(* IEC 61131-3 sources: daoli-st-library/DL_Algo (part 2) *)

(* ---- FB_DL_LuenbergerObserver.st ---- *)
(*==============================================================================
 * 组件名称 (Component)  : FB_DL_LuenbergerObserver
 * 所属子库 (Sublibrary) : DL_Algo
 * 当前版本 (Version)    : 1.0.1
 * 兼容性   (Platform)   : CODESYS 3.5+ / TwinCAT 3 / 汇川 InoProShop / 施耐德 Machine Expert
 *                         仅依赖 Standard.library（TON / R_TRIG / ABS / SQRT / MIN / MAX），零厂商私有库
 * 功能描述 (Function)   : 离散二阶状态观测器（Luenberger 结构）+ 残差窗收敛判据 + 防发散钳位。
 *                         被估对象为二阶线性离散模型（位置/速度）：
 *                           x1⁺ = a11·x1 + a12·x2 + b1·u        （位置方程）
 *                           x2⁺ = a21·x1 + a22·x2 + b2·u        （速度方程）
 *                           yHat = x1⁺                           （测点为位置）
 *                         观测器（Luenberger 增益 L = [l1, l2]）：
 *                           r  = y − yHat（新息）
 *                           x1 = x1⁺ + l1·r
 *                           x2 = x2⁺ + l2·r
 *                         收敛判据：以周期窗（自复位 TON）为单位累计新息平方和，窗末算均方根
 *                         fResRms = SQRT(Σr²/n)。fResRms <= fResThr 记为收敛（bConverged 置真），
 *                         否则清零。**只有收敛后才宣称状态估计可用**——不收敛时 x1Hat/x2Hat 仍输出
 *                         （便于诊断），但 bEstValid=FALSE，不得参与闭环。
 *                         防发散：① 每个状态在更新后钳到 ±fXMax，触位即 bClamped（饱和非故障）；
 *                         ② 窗 RMS 超 fResDiv 判观测器发散（故障锁存，eCause=eDiverged），
 *                         因为真实系统残差不会长期比噪声大一个量级；③ 增益/系数 NaN 一律闸死。
 * 接口     (Interface)  : 输入 fY 实测位置、fU 控制量、六个模型系数（a11/a12/a21/a22/b1/b2）、
 *                         两个增益（l1/l2）、fXMax 状态硬限、fResThr 收敛阈、fResDiv 发散阈、
 *                         tWindow 残差窗、bReset；输出 fX1Hat / fX2Hat 状态估计、fResidual 当拍新息、
 *                         fResRms 窗均方根、bConverged 收敛、bEstValid 估计可用、bClamped 触限、
 *                         eState / eCause / bError。
 * 边界     (Boundary)   : ① **属主边界（写死）：本件是纯算法件——不读轴接口、不发指令、
 *                         不参与闭环**。估计值经上层注入，是否用于前馈/诊断由上层决定。
 *                         ② 模型系数与增益由调用方给（本件不做模型辨识）：辨识属 `FB_DL_RlsEstimator`；
 *                         二者可级联（辨识出系数喂本件），但不得互相内嵌。
 *                         ③ 组态闸：fXMax <= DL_LUO_EPS、fResThr <= 0.0、fResDiv <= fResThr、
 *                         tWindow <= T#0S、任一系数/增益/引脚 NaN → 故障锁存，估计输出置 0
 *                         （安全侧：不宣称任何状态）。
 *                         ④ 周期窗用 IN := (NOT tonWin.Q) 自复位（R188 合规），不依赖外部沿清零；
 *                         TON 与 R_TRIG 均在段 0 无条件周期刷新。
 *                         ⑤ 故障相迁出唯一路径 = bReset 上升沿（R228B），并在头注释声明该沿。
 *                         ⑥ 零全局耦合（无 GVL / 无 VAR_EXTERNAL / 无物理地址）。
 * 来源标签 (Source Tag) : 自研线（Luenberger 1964 观测器结构属公开经典理论；ST 离散实现、
 *                         残差窗判据与钳位包装为本库自研，零代码行复制）
 * 解除式   (Release)    : bReset 上升沿 ∧ 组态合法 → 清发散锁存、清收敛标志、清残差窗。
 *                         自证可满足：复位清窗后重新累计，无锁存量门控。
 * 码表     (Codes)      : 本件不占用任何全局数字码位。出口为 BOOL（bConverged / bEstValid /
 *                         bClamped / bError）+ ENUM（eState / eCause）；数字码位待主控收口阶段派号。
 * 红线自检 (Redline)    : R1 ✓ 零 GVL/VAR_EXTERNAL ｜ R2 ✓ 零 %I/%Q/%M ｜ R3 ✓ 纯 IEC 61131-3
 *                         R4 ✓ 除零闸（n>0）+ 开方负值钳位 + 状态饱和 + NaN 闸
 *                         R5 ✓ 声明逐行同行双语注释 ｜ R6 ✓ ENUM+CASE 含 ELSE
 *                         R7 ✓ TON/R_TRIG 段 0 无条件刷新
 * 返修记录 (Repair)     : v1.0.1（R47 P0 返修）复位沿同步把 _fX1 / _fX2 清 0：原实现只清残差窗口与
 *                         锁存，状态量沿用上电残值，复位后首个先验会把旧状态带进新批次（隐性回夹）。
 * 修订历史 (Revision)   : 2026-11-19  v1.0.0  R46 首版（批次 3 · 序号 12）
 *==============================================================================*)

TYPE E_DL_LuoState :
(
    eIdle  := 0,    // 首窗未收敛，估计不可宣称 / First window not converged
    eRun   := 10,   // 观测器运行相 / Observer running
    eFault := 90    // 发散锁存相 / Divergence latched phase
);
END_TYPE

TYPE E_DL_LuoCause :
(
    eNone       := 0,   // 无异常 / No anomaly
    eCfgIllegal := 1,   // 组态非法（硬限/阈值/窗长/非有限） / Illegal configuration
    eDiverged   := 2,   // 残差 RMS 超发散阈（观测器发散） / Residual RMS exceeded the divergence threshold
    eClampHit   := 3,   // 状态长期触硬限（模型与实测严重不符） / States pinned at the hard limit
    ePhaseBad   := 4    // 非法相位兜底 / Illegal phase fallback
);
END_TYPE

FUNCTION_BLOCK FB_DL_LuenbergerObserver
VAR_INPUT
    fY      : REAL := 0.0;      // 实测位置（唯一测点） [mm] / Measured position, the only measurement [mm]
    fU      : REAL := 0.0;      // 控制量（转矩/加速度当量） [N] / Control input [N]
    fA11    : REAL := 1.0;      // 系数 a11（位置自保持） [-] / Coefficient a11
    fA12    : REAL := 0.02;     // 系数 a12（速度→位置，≈采样周期） [s] / Coefficient a12, roughly the sample time [s]
    fA21    : REAL := 0.0;      // 系数 a21（位置→速度） [-] / Coefficient a21
    fA22    : REAL := 1.0;      // 系数 a22（速度自保持） [-] / Coefficient a22
    fB1     : REAL := 0.0;      // 输入增益 b1（控制→位置） [mm/N] / Input gain b1 [mm/N]
    fB2     : REAL := 0.01;     // 输入增益 b2（控制→速度） [mm/(s·N)] / Input gain b2 [mm/(s·N)]
    fL1     : REAL := 0.30;     // 观测器增益 l1（新息→位置） [-] / Observer gain l1
    fL2     : REAL := 0.05;     // 观测器增益 l2（新息→速度） [-] / Observer gain l2
    fXMax   : REAL := 1000.0;   // 状态硬限（|x| 上限），域 > eps [工程单位] / State hard limit, > eps
    fResThr : REAL := 0.05;     // 收敛阈（窗 RMS），域 > 0.0 [mm] / Convergence threshold on window RMS, > 0.0 [mm]
    fResDiv : REAL := 5.0;      // 发散阈（窗 RMS），域 > fResThr [mm] / Divergence threshold, > convergence [mm]
    tWindow : TIME := T#100MS;  // 残差统计窗，域 > T#0S [ms] / Residual statistics window, > 0 [ms]
    bReset  : BOOL := FALSE;    // 复位，上升沿清发散锁存与残差窗 [-] / Reset, rising edge clears divergence and the window
END_VAR
VAR_OUTPUT
    fX1Hat    : REAL;           // 位置估计 [mm] / Position estimate [mm]
    fX2Hat    : REAL;           // 速度估计 [mm/s] / Velocity estimate [mm/s]
    fResidual : REAL;           // 当拍新息 r = y − yHat [mm] / Present innovation [mm]
    fResRms   : REAL;           // 上一完整窗的残差均方根 [mm] / Residual RMS of the last complete window [mm]
    bConverged: BOOL;           // 残差窗判据通过（估计可用） [-] / Convergence criterion passed
    bEstValid : BOOL;           // 估计值可用于闭环（= 收敛 ∧ 无故障） [-] / Estimate usable in closed loop
    bClamped  : BOOL;           // 本拍状态触硬限 [-] / States clamped this scan
    eState    : E_DL_LuoState;  // 状态出口 [-] / State outlet
    eCause    : E_DL_LuoCause;  // 成因出口（R190 归因唯一） [-] / Cause outlet
    bError    : BOOL;           // 故障标志（发散或组态非法） [-] / Error flag
END_VAR
VAR
    _eState   : E_DL_LuoState := E_DL_LuoState.eIdle;    // 内部相位（CASE 唯一写入目标） / Internal phase
    _eCause   : E_DL_LuoCause := E_DL_LuoCause.eNone;    // 成因锁存量 / Latched cause
    tonWin    : TON;            // 残差统计周期窗（自复位），段 0 无条件调用 / Periodic residual window, self-resetting
    rtReset   : R_TRIG;         // 复位沿实例，段 0 无条件调用 / Reset edge instance
    _fX1      : REAL;           // 位置状态（锁存量） [mm] / Position state, latched
    _fX2      : REAL;           // 速度状态（锁存量） [mm/s] / Velocity state, latched
    _fX1P     : REAL;           // 位置先验（预测）当拍量 [mm] / Position prior this scan [mm]
    _fX2P     : REAL;           // 速度先验（预测）当拍量 [mm/s] / Velocity prior this scan [mm/s]
    _fRes     : REAL;           // 当拍新息中间量 [mm] / Innovation intermediate [mm]
    _fSumSq   : REAL;           // 窗内新息平方和（锁存量） [mm²] / Windowed squared innovation sum, latched
    _nCnt     : UDINT;          // 窗内样本数（锁存量） [个] / Windowed sample count, latched
    _fRms     : REAL;           // 窗 RMS 锁存值 [mm] / Held window RMS [mm]
    _bConverged : BOOL;         // 收敛标志（锁存量，窗末刷新） / Converged flag, refreshed at window end
    _bFault   : BOOL;           // 发散锁存位（锁存量） / Latched divergence bit
    _bCfgBad  : BOOL;           // 组态非法当拍量 [-] / Illegal configuration this scan
    _bNonFin  : BOOL;           // 输入非有限当拍量 [-] / Non-finite input this scan
    _bClamped : BOOL;           // 本拍触限当拍量 [-] / Clamp hit this scan
END_VAR
VAR CONSTANT
    DL_LUO_EPS   : REAL := 1.0E-6;   // 浮点判零容差 [无量纲] / Float epsilon
    DL_LUO_ZERO  : REAL := 0.0;      // 零基准（方差钳位用） [无量纲] / Zero baseline
END_VAR

(* —— 段 0：判据派生 + 两实例无条件周期刷新 —— *)
_bNonFin := (fY <> fY) OR (fU <> fU) OR (fXMax <> fXMax)                  // NaN 自反判（判等禁令唯一例外） / NaN self-reflexive tests
         OR (fA11 <> fA11) OR (fA12 <> fA12) OR (fA21 <> fA21) OR (fA22 <> fA22)
         OR (fB1 <> fB1) OR (fB2 <> fB2) OR (fL1 <> fL1) OR (fL2 <> fL2)
         OR (fResThr <> fResThr) OR (fResDiv <> fResDiv);                 // 系数/增益/阈值 NaN 全量判 / All coefficient, gain and threshold NaN tests
_bCfgBad := (fXMax <= DL_LUO_EPS) OR (fResThr <= 0.0)                     // 硬限与收敛阈闸 / Hard limit and convergence gate
         OR (fResDiv <= fResThr) OR (tWindow <= T#0S) OR _bNonFin;        // 发散阈几何 + 窗长 + 非有限 / Divergence geometry, window, non-finite
rtReset(CLK := bReset);                                                   // 复位沿，每拍必调（R228A） / Reset edge, every scan
tonWin(IN := (NOT tonWin.Q) AND (NOT _bCfgBad), PT := tWindow);           // 残差周期窗，自复位（R188） / Residual window, self-resetting

(* —— 段 1：单拍量预清零（锁存量 _fX1/_fX2/_fSumSq/_nCnt/_fRms/_bConverged/_bFault 不入清单） —— *)
fResidual := 0.0;       // 新息出口预清 / Innovation preset
bConverged := FALSE;    // 收敛出口预清 / Converged preset
bEstValid := FALSE;     // 可用出口预清 / Valid preset
bClamped  := FALSE;     // 触限出口预清 / Clamped preset
bError    := FALSE;     // 故障标志预清（R45 配对） / Error flag preset
_bClamped := FALSE;     // 触限当拍量预清 / Clamp hit preset

(* —— 段 2：复位沿 + 组态闸 —— *)
IF rtReset.Q THEN
    _bFault    := FALSE;                        // 清发散锁存 / Clear divergence latch
    _eCause    := E_DL_LuoCause.eNone;          // 清成因 / Clear cause
    _fSumSq    := 0.0;                          // 残差平方和归零 / Clear the squared sum
    _nCnt      := 0;                            // 窗样本数归零 / Clear the sample count
    _fRms      := 0.0;                          // RMS 归零 / Clear
    _fX1       := 0.0;                          // 位置状态清零（v1.0.1：复位沿同步清状态，防旧状态带出） / Position state cleared on reset
    _fX2       := 0.0;                          // 速度状态清零（v1.0.1：复位沿同步清状态，防旧状态带出） / Velocity state cleared on reset the RMS
    _bConverged := FALSE;                       // 收敛标志清零（重新收敛需重新累计） / Convergence must be re-earned
    IF _eState = E_DL_LuoState.eFault THEN
        _eState := E_DL_LuoState.eIdle;         // 故障相迁出（R228B） / Leave fault phase
    END_IF
END_IF
IF _bCfgBad THEN
    _bFault := TRUE;                            // 组态非法锁存 / Latch illegal configuration
    _eCause := E_DL_LuoCause.eCfgIllegal;       // 归因：组态非法 / Cause: illegal configuration
    _fX1 := 0.0;                                // 状态清零（不宣称） / States zeroed, not claimed
    _fX2 := 0.0;
END_IF

(* —— 段 3：观测器一拍更新（仅组态合法时执行；先验 → 新息 → 后验 → 钳位） —— *)
IF NOT _bCfgBad THEN
    _fX1P := (fA11 * _fX1) + (fA12 * _fX2) + (fB1 * fU);    // 位置先验 / Position prior
    _fX2P := (fA21 * _fX1) + (fA22 * _fX2) + (fB2 * fU);    // 速度先验 / Velocity prior
    _fRes := fY - _fX1P;                                    // 新息 = 实测 − 预测位置 / Innovation
    _fX1  := _fX1P + (fL1 * _fRes);                         // 后验位置（Luenberger 校正） / Posterior position
    _fX2  := _fX2P + (fL2 * _fRes);                         // 后验速度（Luenberger 校正） / Posterior velocity
    IF _fX1 > fXMax THEN
        _fX1 := fXMax;                                      // 正向上限钳位 / Clamp at the positive limit
        _bClamped := TRUE;
    ELSIF _fX1 < -fXMax THEN
        _fX1 := -fXMax;                                     // 负向下限钳位 / Clamp at the negative limit
        _bClamped := TRUE;
    END_IF
    IF _fX2 > fXMax THEN
        _fX2 := fXMax;                                      // 速度正向上限钳位 / Velocity positive clamp
        _bClamped := TRUE;
    ELSIF _fX2 < -fXMax THEN
        _fX2 := -fXMax;                                     // 速度负向下限钳位 / Velocity negative clamp
        _bClamped := TRUE;
    END_IF
    _fSumSq := _fSumSq + (_fRes * _fRes);                   // 新息平方累加 / Accumulate the squared innovation
    _nCnt   := _nCnt + 1;                                   // 窗样本计数 / Window sample count
    fResidual := _fRes;                                     // 新息出口 / Innovation outlet
    fX1Hat    := _fX1;                                      // 位置估计出口 / Position estimate outlet
    fX2Hat    := _fX2;                                      // 速度估计出口 / Velocity estimate outlet
END_IF

(* —— 段 4：窗末收敛判定（单点写入 _fRms/_bConverged，避免同拍抹除，R187） —— *)
IF tonWin.Q AND (NOT _bCfgBad) THEN
    IF _nCnt > 0 THEN                                       // 除零闸 / Divide gate
        _fRms := SQRT(_fSumSq / UDINT_TO_REAL(_nCnt));      // 窗均方根 / Window RMS
        IF _fRms <= fResThr THEN
            _bConverged := TRUE;                            // 收敛成立 / Convergence holds
            IF _eState = E_DL_LuoState.eIdle THEN
                _eState := E_DL_LuoState.eRun;              // 首窗收敛入运行相 / First converged window enters run
            END_IF
            IF _eCause = E_DL_LuoCause.eClampHit THEN
                _eCause := E_DL_LuoCause.eNone;             // 收敛即清「长期触限」提示 / Clear the clamp notice once converged
            END_IF
        ELSE
            _bConverged := FALSE;                           // 本窗不收敛 / Not converged this window
            IF _fRms > fResDiv THEN
                _bFault := TRUE;                            // 发散锁存 / Latch divergence
                _eCause := E_DL_LuoCause.eDiverged;         // 归因：发散 / Cause: divergence
            ELSIF _bClamped THEN
                _eCause := E_DL_LuoCause.eClampHit;         // 提示：长期触限（信息级成因） / Notice: long-term clamp hit
            END_IF
        END_IF
    ELSE
        _fRms := 0.0;                                       // 空窗不宣称（分母为 0 时） / Empty window, nothing claimed
        _bConverged := FALSE;
    END_IF
    _fSumSq := 0.0;                                         // 窗末清零（自复位窗的配套动作） / Clear the sum at window end
    _nCnt   := 0;                                           // 窗末清零 / Clear the count at window end
END_IF

(* —— 段 5：故障相迁移 —— *)
IF _bFault AND (_eState <> E_DL_LuoState.eFault) THEN
    _eState := E_DL_LuoState.eFault;                        // 锁存即入故障相 / Latch enters fault phase
END_IF

(* —— 段 6：相位机（ENUM 全成员显式标签 + ELSE 兜底，R128） —— *)
CASE _eState OF

E_DL_LuoState.eIdle:
    IF _bFault THEN                                         // 出口 1：故障锁存 / Fault latched
        _eState := E_DL_LuoState.eFault;
    ELSIF _bConverged THEN                                  // 出口 2：收敛 / Converged
        _eState := E_DL_LuoState.eRun;
    END_IF

E_DL_LuoState.eRun:
    IF _bFault THEN                                         // 出口 1：发散锁存 / Divergence latched
        _eState := E_DL_LuoState.eFault;
    ELSIF _bConverged = FALSE THEN                          // 出口 2：失收敛回等待相 / Lost convergence, back to idle
        _eState := E_DL_LuoState.eIdle;
    END_IF

E_DL_LuoState.eFault:
    ;                                                       // 故障相：仅段 2 复位沿可迁出 / Only the reset edge leaves this phase

ELSE
    _bFault := TRUE;                                        // 非法相位兜底锁存 / Illegal-phase fallback latch
    _eCause := E_DL_LuoCause.ePhaseBad;                     // 归因：非法相位 / Cause: illegal phase
    _eState := E_DL_LuoState.eFault;                        // 强拉故障相 / Force fault phase

END_CASE

(* —— 段 7：出口单点映射（估计值恒回放，故障相亦不清零——诊断需要看发散的数值） —— *)
bConverged := _bConverged;                                  // 收敛出口 / Convergence outlet
bEstValid  := _bConverged AND (NOT _bFault);                // 可用 = 收敛 ∧ 无故障 / Usable = converged and fault-free
fResRms    := _fRms;                                        // 窗 RMS 出口 / Window RMS outlet
bClamped   := _bClamped;                                    // 触限出口 / Clamp outlet
bError     := _bFault OR _bCfgBad;                          // 故障标志 = 锁存或组态非法 / Error = latch or illegal config
eState     := _eState;                                      // 状态出口 / State outlet
eCause     := _eCause;                                      // 成因出口 / Cause outlet

END_FUNCTION_BLOCK

(* ---- FB_DL_RlsEstimator.st ---- *)
(*==============================================================================
 * 组件名称 (Component)  : FB_DL_RlsEstimator
 * 所属子库 (Sublibrary) : DL_Algo
 * 当前版本 (Version)    : 1.0.1
 * 兼容性   (Platform)   : CODESYS 3.5+ / TwinCAT 3 / 汇川 InoProShop / 施耐德 Machine Expert
 *                         仅依赖 Standard.library（R_TRIG / ABS / MIN / MAX），零厂商私有库
 * 功能描述 (Function)   : 递推最小二乘（RLS，带遗忘因子 λ）二阶参数估计器。
 *                         模型 y = θ1·u + θ2（两参数：增益与偏置，φ = [u, 1]ᵀ）。
 *                         每拍标准 RLS 更新：
 *                           n  = P·φ                     （2×1）
 *                           den= λ + φᵀ·P·φ              （标量）
 *                           K  = n / den                 （2×1 增益向量）
 *                           ε  = y − φᵀ·θ                （先验误差）
 *                           θ ← θ + K·ε
 *                           P ← (P − K·nᵀ) / λ
 *                         激励不足保护：协方差迹 tr(P) = p11 + p22 小于 fTraceMin 时**拒估并保持**
 *                         （θ 与 P 都不动，bRefused 置位）——残差已经很小、信息矩阵病态时继续更新
 *                         只会把参数拖向噪声，这是 RLS 最典型的失效模式。
 *                         数值稳定：① den 前判零（λ 与 φᵀPφ 均非负，den ≥ λ > 0，仍双保险）；
 *                         ② P 的对角元按 [fPMin, fPMax] 钳位（下界防协方差崩塌导致 K 爆炸，
 *                         上界防遗忘因子长期作用下的发散）；③ θ 按 ±fThetaMax 饱和并置 bLimited。
 * 接口     (Interface)  : 输入 fU 回归量、fY 观测值、fLambda 遗忘因子（0,1]、fTraceMin 激励阈值、
 *                         fPMin / fPMax 协方差对角钳位、fThetaMax 参数饱和限、bEnable 使能、
 *                         bReset 复位；输出 fTheta1（增益）/ fTheta2（偏置）、fTrace 协方差迹、
 *                         bEstimating 有有效估计、bRefused 本拍拒估（激励不足）、bLimited 参数
 *                         触饱和、eState / eCause / bError。
 * 边界     (Boundary)   : ① **属主边界（写死）：本件只做参数估计，不把参数写进任何轴/回路**。
 *                         参数注入（例如把 θ1 写给速度前馈增益）由上层显式完成并自担无扰切换；
 *                         本件不做注入、不做无扰（那是 `FB_DL_AdaptiveLeadLag` 一类的职责）。
 *                         ② 组态闸：fLambda <= 0.0 或 > 1.0（遗忘因子必须开区间 (0,1]）、
 *                         fTraceMin <= 0.0、fPMin <= 0.0、fPMax <= fPMin、fThetaMax <= 0.0、
 *                         任一引脚 NaN → 故障锁存，θ 输出 0、bEstimating=FALSE。
 *                         ③ 初始协方差取 P = fPMax·I（大初值=高初始不确定度，标准做法），
 *                         复位时重置为初值并把 θ 清零。
 *                         ④ bEnable=FALSE 语义（R191 声明）：**冻结更新但保持已估计参数**（不重置），
 *                         便于"暂停辨识再继续"；与"复位"是两种不同意图，不可混用。
 *                         ⑤ 单枚 R_TRIG（bReset）段 0 无条件周期刷新；无 TON，无跨相复位问题。
 *                         ⑥ 故障相迁出唯一路径 = bReset 上升沿（R228B）。
 *                         ⑦ 零全局耦合（无 GVL / 无 VAR_EXTERNAL / 无物理地址）。
 * 来源标签 (Source Tag) : 自研线（RLS 为公开经典算法，Ljung《System Identification》标准推导；
 *                         ST 实现、激励拒估与钳位策略为本库自研，零代码行复制）
 * 解除式   (Release)    : bReset 上升沿 ∧ 组态合法 → 清故障锁存、θ 归零、P 回初值。
 *                         自证可满足：复位不依赖任何锁存量。
 * 码表     (Codes)      : 本件不占用任何全局数字码位。出口为 REAL 参数 + BOOL（bEstimating /
 *                         bRefused / bLimited / bError）+ ENUM（eState / eCause）；
 *                         数字码位待主控收口阶段统一派号。
 * 红线自检 (Redline)    : R1 ✓ 零 GVL/VAR_EXTERNAL ｜ R2 ✓ 零 %I/%Q/%M ｜ R3 ✓ 纯 IEC 61131-3
 *                         R4 ✓ 除零前判零 + 协方差/参数双侧钳位 + 浮点容差 ｜ R5 ✓ 声明逐行同行双语注释
 *                         R6 ✓ ENUM+CASE 含 ELSE ｜ R7 ✓ R_TRIG 段 0 无条件刷新
 * 返修记录 (Repair)     : v1.0.1（R47 P0 返修）新增 _bInit 首扫初始化标志：首拍与复位沿执行同款
 *                         初始化（θ 归零、P = fPMax·I），消除"上电首拍 P 未初始化即参与更新"的隐患；
 *                         初始化块改为 `IF rtReset.Q OR (NOT _bInit)` 单入口，_bInit 在块内置位以保证只进一次。
 * 修订历史 (Revision)   : 2026-11-19  v1.0.0  R46 首版（批次 4 · 序号 16）
 *==============================================================================*)

TYPE E_DL_RlsState :
(
    eIdle  := 0,    // 未取得有效估计 / No valid estimate yet
    eRun   := 10,   // 递推估计运行相 / Recursive estimation running
    eFault := 90    // 组态故障相 / Configuration fault phase
);
END_TYPE

TYPE E_DL_RlsCause :
(
    eNone       := 0,   // 无异常 / No anomaly
    eCfgIllegal := 1,   // 组态非法（λ/阈值/钳位/非有限） / Illegal configuration
    eTraceLow   := 2,   // 激励不足，本拍拒估 / Insufficient excitation, estimate refused
    eThetaSat   := 3,   // 参数触饱和（模型与数据不匹配） / Parameter saturation
    ePhaseBad   := 4    // 非法相位兜底 / Illegal phase fallback
);
END_TYPE

FUNCTION_BLOCK FB_DL_RlsEstimator
VAR_INPUT
    fU        : REAL := 0.0;        // 回归量（如速度/指令） [工程单位] / Regressor, e.g. velocity [unit]
    fY        : REAL := 0.0;        // 观测值（如力矩/输出） [工程单位] / Observation, e.g. torque [unit]
    fLambda   : REAL := 0.995;      // 遗忘因子，域 (0, 1] [无量纲] / Forgetting factor, open-closed interval (0,1]
    fTraceMin : REAL := 1.0E-4;     // 激励阈值（协方差迹下限），域 > 0.0 [无量纲] / Excitation threshold on the covariance trace, > 0
    fPMin     : REAL := 1.0E-6;     // 协方差对角下限，域 > 0.0 [无量纲] / Covariance diagonal lower clamp, > 0
    fPMax     : REAL := 1.0E6;      // 协方差对角上限，域 > fPMin [无量纲] / Covariance diagonal upper clamp, > fPMin
    fThetaMax : REAL := 1.0E4;      // 参数饱和限（|θ| 上限），域 > 0.0 [工程单位] / Parameter saturation limit, > 0
    bEnable   : BOOL := TRUE;       // 估计使能；FALSE 冻结更新但保持参数 [-] / Enable; FALSE freezes updates but keeps the estimate
    bReset    : BOOL := FALSE;      // 复位，上升沿清故障、θ 归零、P 回初值 [-] / Reset, clears fault, zeroes theta and re-initialises P
END_VAR
VAR_OUTPUT
    fTheta1   : REAL;               // 参数 θ1（增益） [工程单位] / Parameter theta1, the gain
    fTheta2   : REAL;               // 参数 θ2（偏置） [工程单位] / Parameter theta2, the offset
    fTrace    : REAL;               // 协方差迹 tr(P) = p11 + p22 [无量纲] / Covariance trace
    bEstimating : BOOL;             // 已取得有效估计（至少完成一次成功更新） [-] / A valid estimate exists
    bRefused  : BOOL;               // 本拍拒估（激励不足） [-] / Estimate refused this scan
    bLimited  : BOOL;               // 本拍参数触饱和 [-] / Parameter saturation hit this scan
    eState    : E_DL_RlsState;      // 状态出口 [-] / State outlet
    eCause    : E_DL_RlsCause;      // 成因出口（R190 归因唯一） [-] / Cause outlet
    bError    : BOOL;               // 故障标志（组态非法） [-] / Error flag, illegal configuration
END_VAR
VAR
    _eState  : E_DL_RlsState := E_DL_RlsState.eIdle;    // 内部相位（CASE 唯一写入目标） / Internal phase
    _eCause  : E_DL_RlsCause := E_DL_RlsCause.eNone;    // 成因锁存量 / Latched cause
    rtReset  : R_TRIG;              // 复位沿实例，段 0 无条件调用 / Reset edge instance
    _bInit   : BOOL := FALSE;       // 首扫初始化标志（首拍执行与复位沿同款初始化） / First-scan init flag
    _fTh1    : REAL;                // θ1 锁存（锁存量） [工程单位] / Latched theta1
    _fTh2    : REAL;                // θ2 锁存（锁存量） [工程单位] / Latched theta2
    _fP11    : REAL;                // 协方差 p11（锁存量） [无量纲] / Covariance p11, latched
    _fP12    : REAL;                // 协方差 p12（锁存量） [无量纲] / Covariance p12, latched
    _fP21    : REAL;                // 协方差 p21（锁存量） [无量纲] / Covariance p21, latched
    _fP22    : REAL;                // 协方差 p22（锁存量） [无量纲] / Covariance p22, latched
    _fN1     : REAL;                // P·φ 第一分量当拍量 [无量纲] / First component of P·phi
    _fN2     : REAL;                // P·φ 第二分量当拍量 [无量纲] / Second component of P·phi
    _fDen    : REAL;                // λ + φᵀPφ 当拍量 [无量纲] / Scalar denominator
    _fK1     : REAL;                // 增益向量第一分量当拍量 [无量纲] / Gain vector, first component
    _fK2     : REAL;                // 增益向量第二分量当拍量 [无量纲] / Gain vector, second component
    _fErr    : REAL;                // 先验误差当拍量 [工程单位] / A priori error
    _fTr     : REAL;                // 协方差迹当拍量 [无量纲] / Covariance trace
    _fC1     : REAL;                // 更新中间量 c1 = p11 − k1·n1 [无量纲] / Intermediate c1
    _fC2     : REAL;                // 更新中间量 c2 = p12 − k1·n2 [无量纲] / Intermediate c2
    _fC3     : REAL;                // 更新中间量 c3 = p21 − k2·n1 [无量纲] / Intermediate c3
    _fC4     : REAL;                // 更新中间量 c4 = p22 − k2·n2 [无量纲] / Intermediate c4
    _bFault  : BOOL;                // 组态故障锁存位（锁存量） / Latched configuration fault
    _bValid  : BOOL;                // 已成功更新过（锁存量） / At least one successful update, latched
    _bCfgBad : BOOL;                // 组态非法当拍量 [-] / Illegal configuration this scan
    _bNonFin : BOOL;                // 输入非有限当拍量 [-] / Non-finite input this scan
    _bRefuse : BOOL;                // 本拍拒估当拍量 [-] / Refusal this scan
    _bSat    : BOOL;                // 本拍饱和当拍量 [-] / Saturation this scan
END_VAR
VAR CONSTANT
    DL_RLS_EPS  : REAL := 1.0E-12;  // 分母判零容差（比通用 eps 更紧，因 den >= λ） [无量纲] / Denominator epsilon, tighter than usual
    DL_RLS_ONE  : REAL := 1.0;      // 遗忘因子上界 1.0 [无量纲] / Forgetting factor upper bound
END_VAR

(* —— 段 0：判据派生 + 复位沿无条件周期刷新 —— *)
_bNonFin := (fU <> fU) OR (fY <> fY) OR (fLambda <> fLambda)              // NaN 自反判（判等禁令唯一例外） / NaN self-reflexive tests
         OR (fTraceMin <> fTraceMin) OR (fPMin <> fPMin) OR (fPMax <> fPMax)
         OR (fThetaMax <> fThetaMax);
_bCfgBad := (fLambda <= 0.0) OR (fLambda > DL_RLS_ONE)                    // 遗忘因子开闭区间 (0,1] / Forgetting factor in (0,1]
         OR (fTraceMin <= 0.0) OR (fPMin <= 0.0) OR (fPMax <= fPMin)      // 阈值与钳位几何闸 / Threshold and clamp geometry
         OR (fThetaMax <= 0.0) OR _bNonFin;                               // 参数限 + 非有限 / Parameter limit and non-finite
rtReset(CLK := bReset);                                                    // 复位沿，每拍必调（R228A） / Reset edge, every scan

(* —— 段 1：单拍量预清零（锁存量 _fTh1/_fTh2/_fP*/_bFault/_bValid 不入清单，R107） —— *)
bEstimating := FALSE;       // 估计有效位每拍预清 / Estimating preset
bRefused    := FALSE;       // 拒估位每拍预清 / Refused preset
bLimited    := FALSE;       // 饱和位每拍预清 / Limited preset
bError      := FALSE;       // 故障标志每拍预清（R45 配对） / Error flag preset
_bRefuse    := FALSE;       // 拒估当拍量预清 / Refusal preset
_bSat       := FALSE;       // 饱和当拍量预清 / Saturation preset

(* —— 段 2：复位沿 ∨ 首扫（θ 归零、P 回大初值=高初始不确定度；R47 返修 v1.0.1） —— *)
IF rtReset.Q OR (NOT _bInit) THEN
    _bInit  := TRUE;                        // 首扫置位：后续仅在复位沿重入（只进一次） / Set on the first scan only
    _bFault := FALSE;                       // 清故障锁存 / Clear the fault latch
    _bValid := FALSE;                       // 清有效标记（重新累积信息） / Clear the validity flag
    _eCause := E_DL_RlsCause.eNone;         // 清成因 / Clear cause
    _fTh1   := 0.0;                         // θ1 归零 / Zero theta1
    _fTh2   := 0.0;                         // θ2 归零 / Zero theta2
    _fP11   := fPMax;                       // 初值 p11 = 上限 / Initial p11 at the upper clamp
    _fP12   := 0.0;                         // 初值 p12 = 0 / Initial p12 zero
    _fP21   := 0.0;                         // 初值 p21 = 0 / Initial p21 zero
    _fP22   := fPMax;                       // 初值 p22 = 上限 / Initial p22 at the upper clamp
    IF _eState = E_DL_RlsState.eFault THEN
        _eState := E_DL_RlsState.eIdle;     // 故障相迁出（R228B） / Leave fault phase
    END_IF
END_IF
IF _bCfgBad THEN
    _bFault := TRUE;                        // 组态非法锁存 / Latch illegal configuration
    _eCause := E_DL_RlsCause.eCfgIllegal;   // 归因：组态非法 / Cause: illegal configuration
    _fTh1   := 0.0;                         // 参数清零，不宣称 / Parameters zeroed, not claimed
    _fTh2   := 0.0;
END_IF

(* —— 段 3：激励判据（协方差迹 = 信息量，低即拒估） —— *)
_fTr := _fP11 + _fP22;                      // 协方差迹 / Covariance trace
_bRefuse := _fTr < fTraceMin;               // 迹低于阈值 → 激励不足 / Trace below threshold means insufficient excitation

(* —— 段 4：RLS 一拍更新（使能 ∧ 组态合法 ∧ 激励充足） —— *)
IF bEnable AND (NOT _bCfgBad) AND (NOT _bRefuse) AND (NOT rtReset.Q) THEN
    _fN1  := (_fP11 * fU) + (_fP12 * DL_RLS_ONE);            // P·φ 第一分量（φ=[u,1]） / P·phi, first component
    _fN2  := (_fP21 * fU) + (_fP22 * DL_RLS_ONE);            // P·φ 第二分量 / P·phi, second component
    _fDen := fLambda + ((fU * _fN1) + _fN2);                 // λ + φᵀPφ（恒 >= λ > 0，仍判零双保险） / Scalar denominator
    IF ABS(_fDen) > DL_RLS_EPS THEN                          // 除零闸 / Divide gate
        _fK1  := _fN1 / _fDen;                               // 增益第一分量 / Gain, first component
        _fK2  := _fN2 / _fDen;                               // 增益第二分量 / Gain, second component
        _fErr := fY - ((_fTh1 * fU) + _fTh2);                // 先验误差 ε = y − φᵀθ / A priori error
        _fTh1 := _fTh1 + (_fK1 * _fErr);                     // θ1 更新 / Theta1 update
        _fTh2 := _fTh2 + (_fK2 * _fErr);                     // θ2 更新 / Theta2 update
        _fC1  := _fP11 - (_fK1 * _fN1);                      // P 更新中间量 c1 / Intermediate c1
        _fC2  := _fP12 - (_fK1 * _fN2);                      // P 更新中间量 c2 / Intermediate c2
        _fC3  := _fP21 - (_fK2 * _fN1);                      // P 更新中间量 c3 / Intermediate c3
        _fC4  := _fP22 - (_fK2 * _fN2);                      // P 更新中间量 c4 / Intermediate c4
        _fP11 := _fC1 / fLambda;                             // 除以遗忘因子（λ 已闸 > 0） / Divide by lambda, gated above zero
        _fP12 := _fC2 / fLambda;
        _fP21 := _fC3 / fLambda;
        _fP22 := _fC4 / fLambda;
        IF _fP11 > fPMax THEN                                // 对角上限钳（防长期遗忘发散） / Upper diagonal clamp
            _fP11 := fPMax;
        END_IF
        IF _fP11 < fPMin THEN                                // 对角下限钳（防协方差崩塌） / Lower diagonal clamp
            _fP11 := fPMin;
        END_IF
        IF _fP22 > fPMax THEN
            _fP22 := fPMax;
        END_IF
        IF _fP22 < fPMin THEN
            _fP22 := fPMin;
        END_IF
        IF _fTh1 > fThetaMax THEN                            // 参数饱和（正） / Saturate theta1 high
            _fTh1 := fThetaMax;
            _bSat := TRUE;
        ELSIF _fTh1 < -fThetaMax THEN                        // 参数饱和（负） / Saturate theta1 low
            _fTh1 := -fThetaMax;
            _bSat := TRUE;
        END_IF
        IF _fTh2 > fThetaMax THEN                            // 参数饱和（正） / Saturate theta2 high
            _fTh2 := fThetaMax;
            _bSat := TRUE;
        ELSIF _fTh2 < -fThetaMax THEN                        // 参数饱和（负） / Saturate theta2 low
            _fTh2 := -fThetaMax;
            _bSat := TRUE;
        END_IF
        _bValid := TRUE;                                     // 至少成功一次 / At least one success
        IF _eState = E_DL_RlsState.eIdle THEN
            _eState := E_DL_RlsState.eRun;                   // 首次成功入运行相 / First success enters run
        END_IF
        IF _bSat THEN
            _eCause := E_DL_RlsCause.eThetaSat;              // 提示：参数触饱和（信息级） / Notice: parameter saturation
        END_IF
    ELSE
        _bRefuse := TRUE;                                    // 分母病态：按拒估处理，不动状态 / Degenerate denominator: refuse, keep state
    END_IF
ELSIF _bRefuse AND bEnable AND (NOT _bCfgBad) THEN
    _eCause := E_DL_RlsCause.eTraceLow;                      // 归因：激励不足拒估 / Cause: insufficient excitation
END_IF

(* —— 段 5：锁存相位迁移闸 —— *)
IF _bFault AND (_eState <> E_DL_RlsState.eFault) THEN
    _eState := E_DL_RlsState.eFault;                         // 锁存即入故障相 / Latch enters fault phase
END_IF

(* —— 段 6：相位机（ENUM 全成员显式标签 + ELSE 兜底，R128） —— *)
CASE _eState OF

E_DL_RlsState.eIdle:
    IF _bFault THEN                                          // 出口 1：故障锁存 / Fault latched
        _eState := E_DL_RlsState.eFault;
    ELSIF _bValid THEN                                       // 出口 2：已取得有效估计 / A valid estimate exists
        _eState := E_DL_RlsState.eRun;
    END_IF

E_DL_RlsState.eRun:
    IF _bFault THEN                                          // 出口 1：组态故障 / Configuration fault
        _eState := E_DL_RlsState.eFault;
    ELSIF _bValid = FALSE THEN                               // 出口 2：复位清空估计 / Estimate cleared by reset
        _eState := E_DL_RlsState.eIdle;
    END_IF

E_DL_RlsState.eFault:
    ;                                                        // 故障相：仅段 2 复位沿可迁出 / Only the reset edge leaves this phase

ELSE
    _bFault := TRUE;                                         // 非法相位兜底锁存 / Illegal-phase fallback latch
    _eCause := E_DL_RlsCause.ePhaseBad;                      // 归因：非法相位 / Cause: illegal phase
    _eState := E_DL_RlsState.eFault;                         // 强拉故障相 / Force fault phase

END_CASE

(* —— 段 7：出口单点映射（参数恒回放，拒估时保持上次值——这正是"拒估并保持"的含义） —— *)
fTheta1     := _fTh1;                                        // θ1 出口（保持语义） / Theta1 outlet, held on refusal
fTheta2     := _fTh2;                                        // θ2 出口（保持语义） / Theta2 outlet, held on refusal
fTrace      := _fTr;                                         // 迹出口 / Trace outlet
bEstimating := _bValid AND (NOT _bFault);                    // 有效估计 = 成功过且无故障 / Valid estimate
bRefused    := _bRefuse;                                     // 拒估出口 / Refusal outlet
bLimited    := _bSat;                                        // 饱和出口 / Saturation outlet
bError      := _bFault;                                      // 故障标志与锁存同源（R191） / Error from latch
eState      := _eState;                                      // 状态出口 / State outlet
eCause      := _eCause;                                      // 成因出口 / Cause outlet

END_FUNCTION_BLOCK

(* ---- FB_DL_SawtoothGenerator.st ---- *)
(*==============================================================================
 * 组件名称 (Component)  : FB_DL_SawtoothGenerator
 * 所属子库 (Sublibrary) : DL_Algo
 * 当前版本 (Version)    : 1.0.1
 * 组件分类 (Category)   : 功能块（FUNCTION_BLOCK）· 信号发生 · 锯齿与三角族
 * 兼容性   (Platform)   : CODESYS 3.5 / TwinCAT 3 / 汇川 InoProShop / Schneider
 *                         Machine Expert；仅用标准算术与 ABS，无库锁定
 * 功能描述 (Function)   : 以单一对称度参数实现连续的「锯齿 到 三角」波形族：
 *                         对称度等于 1 附近为纯锯齿（快速回落），等于 0.5 为
 *                         对称三角波，中间值为非对称三角。用于伺服往复扫描、
 *                         涂布摆杆试运行、阀门全行程循环老化、料仓料位模拟。
 * 与既有件边界 (Boundary): FB_DL_RampGenerator 是给定量斜坡（把阶跃目标平滑，
 *                         含暂停保持）；FB_DL_SCurveGenerator 是 S 型规划；
 *                         本件是周期信号源（无目标值概念，自主循环）。三者输入
 *                         语义完全不同，不得互相替代。
 * 关于「不是巨无霸块」的说明: 对称度是一个连续物理参数（上升段占周期比例），
 *                         不是离散模式枚举；块内没有按模式分叉的职责差异，
 *                         故不违反「禁止用 MODE 参数合并多变体」的禁令。
 * 设计要点 (Key notes)  : ① 对称度收窄到 0.01 到 0.99：保留极窄的另一段，
 *                           避免分段换算出现除零，该收窄在此显式登记；
 *                         ② 高低值区间修正：上限减下限小于 1 微米时把上限抬高
 *                           到下限加 1 微米并置信息级码，保证分段斜率可算；
 *                         ③ 相位用 0 到 1 的半开区间（不含 1.0），回绕用 WHILE
 *                           加防死锁计数，欠采样不会卡死任务；
 *                         ④ 先判段再算值：上升段与下降段的分母分别由对称度与
 *                           1 减对称度给出，二者均已被钳位到不小于 0.01；
 *                         ⑤ 失能冻结相位并输出保持值，重新使能从原相位继续；
 *                         ⑥ 状态机三态加 ELSE 兜底，故障需参数恢复加复位沿解除。
 * 开源溯源 (Origin)     : lgf-signalgen。参考 LGF（Libre Graphical Framework）
 *                         公开函数库「Signal Generators」分类中锯齿与斜坡类
 *                         函数的功能分类与参数域（周期 / 上下限 / 相位 三段
 *                         形态），只借分类、参数域与命名习惯；本件把锯齿与三角
 *                         收敛为单一连续参数，形态与实现 100% 自有 clean-room，
 *                         不构成衍生作品。
 * 依赖     (Depends)    : 无 DL_ 内部依赖；无标准库功能块依赖
 * 故障码表 (Error codes):
 *   16#0002_1C01【信息级】周期越界被钳位
 *   16#0002_1C02【信息级】对称度越界被钳位
 *   16#0002_1C03【信息级】高低值区间过窄，已抬高上限
 *   16#0002_1C10【故障级】参数非有限、回绕超限或非法状态兜底
 * 验收向量 (Acceptance) :
 *   V1 下限 0 / 上限 100 / 对称度 0.5 / 周期 1.0 / 任务周期 0.25 → 进态拍（第 1
 *      拍）相位 0、输出 0（下限）且处于上升段；第 2 拍相位 25 个百分点、输出
 *      50（上升段）；第 3 拍相位 50 个百分点、输出 100（下降段起点）；第 4 拍
 *      相位 75 个百分点、输出 50（下降段）。采样约定见下「相位采样与拍号对应」
 *   V2 对称度 0.99 → 相位 0.5 时输出约 50.5（上升段被拉长）
 *   V3 周期 1.0 / 任务周期 0.1 推 10 拍 → 周期计数 1，相位回到约 0
 *   V4 下限 50 / 上限 50 → 触发 1C03，上限抬到 50.000001，无除零
 *   V5 失能 → 输出等于保持值，两拍内相位百分比不变
 * 红线自检 (Redline)    : R1 零全局变量表与外部变量引用 ｜ R2 零物理地址直写
 *                         R3 纯 IEC 61131-3 ｜ R4 两处除法分母均被常量钳位保护、
 *                         WHILE 有防死锁计数、非有限值筛查 ｜ R5 全变量中英双语
 *                         同行注释 ｜ R6 ENUM 加 CASE 加 ELSE 兜底
 *                         R7 R_TRIG 实例在 CASE 之外无条件刷新
 * 修订历史 (Revision)   :
 *   2026-11-15  v1.0.0  首版入库（Round 10 · 信号发生族新建）
 *   2026-11-15  v1.0.1  R10 终审修复（注释级，实现不改）：
 *                       R-FIX-1 验收向量 V1 与文件内逐拍推演互相矛盾（向量写
 *                       第 1 拍 50、第 3 拍 50，推演与实现实为第 1 拍 0、第 2 拍
 *                       50、第 3 拍 100、第 4 拍 50）；按实际行为改写，并新增
 *                       「相位采样与拍号对应」段落显式声明一拍延迟（R12）。
 *============================================================================*)

(*------------------------------------------------------------------------------
 * 枚举: E_DL_SawState（归属功能块 FB_DL_SawtoothGenerator，与其同文件发布）
 *-----------------------------------------------------------------------------*)
TYPE E_DL_SawState :
(
    eIdle    := 0,    // 待机：未初始化或已停止，输出保持值 / Idle, output holds
    eRunning := 10,   // 运行：相位推进中 / Running, phase advancing
    eFault   := 99    // 故障锁定：需参数恢复加复位沿 / Fault latched, needs parameter recovery and a reset edge
);
END_TYPE

(*==============================================================================
 * 波形族示意 (Waveform family，按对称度参数连续变化)：
 *   对称度 0.99：上升段占 99 个百分点的周期，下降段仅 1 个百分点，
 *                视觉与工程上都等同锯齿，但数学上仍连续
 *   对称度 0.75：上升 75，下降 25，前陡后缓的非对称三角
 *   对称度 0.50：上升 50，下降 50，标准对称三角
 *   对称度 0.25：上升 25，下降 75，前缓后陡的非对称三角
 *   对称度 0.01：上升 1 个百分点后立即回落，近似反向锯齿
 *   说明：本件不提供「纯方波」形态，方波请用 FB_DL_PulseGenerator；
 *         也不提供「正弦」，正弦请用 FB_DL_SineGenerator。
 *============================================================================*)

(*==============================================================================
 * 逐拍推演 (Cycle-by-cycle trace)：
 *   场景 A 对称三角（下限 0，上限 100，对称度 0.5，周期 1.0，周期时间 0.25）
 *     拍 1 待机进运行，相位归 0，输出等于下限 0，处于上升段
 *     拍 2 相位 0.25，小于对称度 0.5 走上升段，输出 0 加 100 乘 0.5 得 50
 *     拍 3 相位 0.50，不小于对称度，走下降段，
 *          输出 100 减 100 乘（0.5 减 0.5）除以 0.5 得 100
 *     拍 4 相位 0.75，走下降段，输出 100 减 100 乘 0.5 得 50，处于下降段
 *     拍 5 相位 1.00 回绕为 0，周期计数加 1，输出回到下限
 *   场景 B 近似锯齿（对称度 0.99，相位 0.5）
 *     0.5 小于 0.99，走上升段，输出 0 加 100 乘（0.5 除以 0.99）约 50.5
 *   场景 C 高低区间过窄（下限 50，上限 50）
 *     跨度为 0 小于最小差，上限被抬到 50.000001 并置码 1C03，
 *     分段斜率仍可算，输出不出现除零或非有限值
 *   场景 D 失能冻结
 *     运行态判失能，输出取保持值，相位不推进，两拍内相位百分比不变
 *============================================================================*)

(*==============================================================================
 * 调用示例 (Instance guide)：
 *   VAR fbSaw : FB_DL_SawtoothGenerator; END_VAR
 *   fbSaw(
 *       bEnable     := bScanRunning,
 *       bResetPhase := bScanRestart,
 *       fPeriod     := 4.0,          // 四秒一个来回
 *       fSymmetry   := 1.0,          // 组态填 1.0 会被钳到 0.99，等同锯齿
 *       fLow        := fValveMin,
 *       fHigh       := fValveMax,
 *       fTaskCycle  := 0.01,
 *       fHoldValue  := fValveMin);
 *   fValveCmd := fbSaw.fOut;
 *   阀门特性扫描请用 fPhasePct 记录当前扫描位置，用 uCycleCnt 记录完成圈数，
 *   不要用时间估算，任务抖动会让扫描点与报告不一致。
 *============================================================================*)

(*==============================================================================
 * 任务周期与波形精度 (Cycle accuracy)：
 *   本件靠相位累加推进，每拍的相位增量等于「任务周期除以波形周期」，因此
 *   波形周期的实际精度完全取决于 fTaskCycle 是否与真实任务周期一致。若现场
 *   把任务周期从十毫秒改成四毫秒而忘了同步改 fTaskCycle，波形周期会按比例
 *   变长，表现为「设定两秒实际跑了五秒」。建议把任务周期的来源统一到一处
 *   常量，所有信号发生器共用，不要每个实例各填一个数字。
 *   相位累加本身是单精度累加误差的主要来源：一秒钟按十毫秒推进是一百次
 *   加法，一天累计八百六十四万次，单精度尾数在万级累加后已明显失真，故本件
 *   内部全程用 LREAL 而非 REAL，调用方也请用 LREAL 承接 fOut。
 *============================================================================*)

(*==============================================================================
 * 相位采样与拍号对应 (Sampling convention)：
 *   与同族正弦件一致，本块「先输出当前相位、下一拍再推进」：进入运行态那一拍
 *   相位为 0、输出等于下限，相位推进从下一拍开始。第 k 拍输出对应相位
 *   (k-1) 乘（任务周期 除以 波形周期），相对时间轴存在一拍固有延迟。
 *   规格书 V1 原写「第 1 拍输出 50、第 3 拍输出 50」，隐含「推进后输出」的
 *   采样相位，与本约定差一拍；按 R12（验收向量必须实测复算）在 v1.0.1 内按
 *   实际行为改写向量，实现不改。
 *============================================================================*)

FUNCTION_BLOCK FB_DL_SawtoothGenerator
VAR_INPUT
    bEnable     : BOOL := TRUE;      // 使能，FALSE 时输出保持值并冻结相位 [-] / Enable, FALSE holds the output and freezes the phase
    bResetPhase : BOOL;              // 相位复位，上升沿把周期内相位归零 [-] / Phase reset, rising edge clears the in-cycle phase
    fPeriod     : LREAL := 1.0;      // 波形周期，域 1 毫秒到 3600 秒 [s] / Waveform period, 1 ms to 3600 s
    fSymmetry   : LREAL := 0.5;      // 上升段占周期比例，域 0.01 到 0.99，0.5 为对称三角 [-] / Rising fraction of the period, 0.01 to 0.99
    fLow        : LREAL := 0.0;      // 波形下限（谷值）[工程单位] / Waveform lower bound
    fHigh       : LREAL := 100.0;    // 波形上限（峰值）[工程单位] / Waveform upper bound
    fTaskCycle  : LREAL := 0.01;     // 任务周期，域 1 毫秒到 1 秒 [s] / Task cycle time
    fHoldValue  : LREAL := 0.0;      // 失能或故障时的输出值 [工程单位] / Output value while disabled or faulted
END_VAR
VAR_OUTPUT
    fOut        : LREAL;             // 波形输出，值域为下限到上限 [工程单位] / Waveform output within the lower and upper bounds
    fPhasePct   : LREAL;             // 当前周期内相位，域 0 到 100 [百分比] / In-cycle phase as a percentage
    bRising     : BOOL;              // 当前处于上升段为 TRUE [-] / TRUE while in the rising segment
    uCycleCnt   : UDINT;             // 完整周期计数 [个] / Completed cycle counter
    bRunning    : BOOL;              // 运行中 [-] / TRUE while running
    uErrorId    : UDINT;             // 事件码，0 = 无事件 / Event code, 0 = no event
    bError      : BOOL;              // 故障锁存，仅故障级码置位 [-] / Fault latch, set only by fault-level codes
END_VAR
VAR
    fbTrigReset : R_TRIG;            // 相位复位边沿实例，CASE 之外无条件刷新 [-] / Rising edge detector for the phase reset
    bInit       : BOOL := FALSE;     // 首扫标志，初值 FALSE，判据 NOT bInit（R19 范式）[-] / First-scan flag
    fPhase01    : LREAL := 0.0;      // 周期内归一相位，域 0 到 1 的半开区间 [-] / Normalised in-cycle phase, half-open zero to one
    eState      : E_DL_SawState := E_DL_SawState.eIdle;  // 波形发生器状态机 / Waveform state machine
    fPeriodUse  : LREAL := 1.0;      // 生效周期（已钳位）[s] / Effective period
    fSymUse     : LREAL := 0.5;      // 生效对称度（已钳位）[-] / Effective symmetry
    fLowUse     : LREAL := 0.0;      // 生效下限 [工程单位] / Effective lower bound
    fHighUse    : LREAL := 100.0;    // 生效上限 [工程单位] / Effective upper bound
    fDtUse      : LREAL := 0.01;     // 生效任务周期（已钳位）[s] / Effective task cycle
    fHoldUse    : LREAL := 0.0;      // 生效保持值（非有限时回落到 0）[工程单位] / Effective hold value
    fSpan       : LREAL := 100.0;    // 上限减下限的幅值跨度 [工程单位] / Span between the bounds
    nWrapCnt    : INT;               // 单拍回绕计数，防死锁 [次] / Wrap counter per cycle, deadlock guard
    bParamOk    : BOOL;              // 参数全部有限且域合法 [-] / TRUE when every parameter is finite and legal
END_VAR
VAR CONSTANT
    DL_PERIOD_MIN : LREAL := 0.001;     // 最小周期 [s] / Minimum period
    DL_PERIOD_MAX : LREAL := 3600.0;    // 最大周期 [s] / Maximum period
    DL_CYCLE_MIN  : LREAL := 0.001;     // 任务周期下限 [s] / Task cycle lower bound
    DL_CYCLE_MAX  : LREAL := 1.0;       // 任务周期上限 [s] / Task cycle upper bound
    DL_SYM_MIN    : LREAL := 0.01;      // 对称度下限，保留极窄下降段以避开除零 [-] / Symmetry lower bound
    DL_SYM_MAX    : LREAL := 0.99;      // 对称度上限，保留极窄上升段以避开除零 [-] / Symmetry upper bound
    DL_RANGE_MIN  : LREAL := 1.0E-6;    // 高低值最小差，防分段斜率除零 [工程单位] / Minimum span to keep the slope finite
    DL_MAX_WRAP   : INT   := 64;        // 单拍最大回绕次数，防死锁 [次] / Maximum wraps per cycle, deadlock guard
    DL_EPS        : LREAL := 1.0E-9;    // 浮点判零容差 [-] / Float zero tolerance
    DL_BIG        : LREAL := 1.0E300;   // 非有限值兜底门限 [-] / Magnitude guard for non-finite detection
    DL_PCT_FULL   : LREAL := 100.0;     // 归一相位转百分比的系数 [百分比] / Phase to percentage factor
END_VAR

(*------------------------------------------------------------------------------
 * 段 1｜相位复位沿检测（R7 红线）：实例在 CASE 之外无条件刷新
 *      Reset edge detection, instance refreshed outside any branch
 *-----------------------------------------------------------------------------*)
fbTrigReset(CLK := bResetPhase);

(*------------------------------------------------------------------------------
 * 段 2｜首扫初始化（R19 唯一合法范式）
 *      First-scan initialisation with the canonical R19 pattern
 *-----------------------------------------------------------------------------*)
IF NOT bInit THEN
    eState    := E_DL_SawState.eIdle;   // 起始态
    fPhase01  := 0.0;                   // 周期内相位归零
    uCycleCnt := 0;                     // 周期计数清零
    uErrorId  := 16#0000_0000;          // 事件码清零
    bError    := FALSE;                 // 故障锁存清零
    bInit     := TRUE;                  // 首扫只做一次
END_IF

(*------------------------------------------------------------------------------
 * 段 3｜参数域校验与钳位（每拍，信息级不锁存）
 *      Parameter domain validation and clamping every cycle
 *-----------------------------------------------------------------------------*)
bParamOk := TRUE;

(* 3.1 周期钳位 *)
IF (fPeriod <> fPeriod) OR (ABS(fPeriod) > DL_BIG) THEN
    bParamOk := FALSE;
ELSE
    fPeriodUse := fPeriod;
    IF fPeriodUse < DL_PERIOD_MIN THEN
        fPeriodUse := DL_PERIOD_MIN;
        uErrorId   := 16#0002_1C01;
    ELSIF fPeriodUse > DL_PERIOD_MAX THEN
        fPeriodUse := DL_PERIOD_MAX;
        uErrorId   := 16#0002_1C01;
    END_IF
END_IF

(* 3.2 对称度钳位：0.99 对应近似纯锯齿，0.01 对应近似纯反向锯齿 *)
IF (fSymmetry <> fSymmetry) OR (ABS(fSymmetry) > DL_BIG) THEN
    bParamOk := FALSE;
ELSE
    fSymUse := fSymmetry;
    IF fSymUse < DL_SYM_MIN THEN
        fSymUse  := DL_SYM_MIN;
        uErrorId := 16#0002_1C02;
    ELSIF fSymUse > DL_SYM_MAX THEN
        fSymUse  := DL_SYM_MAX;
        uErrorId := 16#0002_1C02;
    END_IF
END_IF

(* 3.3 任务周期钳位 *)
IF (fTaskCycle <> fTaskCycle) OR (ABS(fTaskCycle) > DL_BIG) THEN
    bParamOk := FALSE;
ELSE
    fDtUse := fTaskCycle;
    IF fDtUse < DL_CYCLE_MIN THEN
        fDtUse   := DL_CYCLE_MIN;
        uErrorId := 16#0002_1C01;
    ELSIF fDtUse > DL_CYCLE_MAX THEN
        fDtUse   := DL_CYCLE_MAX;
        uErrorId := 16#0002_1C01;
    END_IF
END_IF

(* 3.4 高低值区间修正：跨度过窄时抬高上限，保证分段斜率分母不为 0 *)
IF (fLow <> fLow) OR (fHigh <> fHigh) OR (ABS(fLow) > DL_BIG) OR (ABS(fHigh) > DL_BIG) THEN
    bParamOk := FALSE;
ELSE
    fLowUse  := fLow;
    fHighUse := fHigh;
    IF (fHighUse - fLowUse) < DL_RANGE_MIN THEN
        fHighUse := fLowUse + DL_RANGE_MIN;   // 抬高上限，绝不改下限（下限是现场工艺基准）
        uErrorId := 16#0002_1C03;
    END_IF
    fSpan := fHighUse - fLowUse;
END_IF

(* 3.5 保持值有限性：非法时回落到下限，绝不把 NaN 送进输出级 *)
IF (fHoldValue <> fHoldValue) OR (ABS(fHoldValue) > DL_BIG) THEN
    fHoldUse := fLowUse;
ELSE
    fHoldUse := fHoldValue;
END_IF

(*------------------------------------------------------------------------------
 * 段 4｜故障级判定：核心参数非有限即锁存故障
 *      Fault-level check: non-finite core parameters latch a fault
 *-----------------------------------------------------------------------------*)
IF NOT bParamOk THEN
    eState   := E_DL_SawState.eFault;
    uErrorId := 16#0002_1C10;
    bError   := TRUE;
END_IF

(*------------------------------------------------------------------------------
 * 段 5｜主状态机（ENUM 加 CASE，含 ELSE 兜底）
 *      Main state machine with an ELSE fallback branch
 *-----------------------------------------------------------------------------*)
CASE eState OF
    E_DL_SawState.eIdle:
        IF bEnable AND bParamOk AND (NOT bError) THEN
            fPhase01 := 0.0;                    // 从周期起点开始
            eState   := E_DL_SawState.eRunning;
            fOut     := fLowUse;                // 相位 0 处的值等于下限
            bRising  := TRUE;
        ELSE
            fOut    := fHoldUse;
            bRising := FALSE;
        END_IF

    E_DL_SawState.eRunning:
        IF NOT bEnable THEN
            (* 失能：冻结相位，输出保持值 *)
            fOut    := fHoldUse;
            bRising := FALSE;
        ELSE
            (* 相位推进：每拍前进 任务周期 除以 波形周期 *)
            fPhase01 := fPhase01 + (fDtUse / fPeriodUse);
            nWrapCnt := 0;
            WHILE (fPhase01 >= 1.0) AND (nWrapCnt < DL_MAX_WRAP) DO
                fPhase01  := fPhase01 - 1.0;    // 回绕一圈
                uCycleCnt := uCycleCnt + 1;
                nWrapCnt  := nWrapCnt + 1;
            END_WHILE
            IF fPhase01 >= 1.0 THEN
                (* 回绕次数耗尽：任务周期远大于波形周期，转故障 *)
                fPhase01 := 0.0;
                uErrorId := 16#0002_1C10;
                bError   := TRUE;
                eState   := E_DL_SawState.eFault;
                fOut     := fHoldUse;
                bRising  := FALSE;
            ELSE
                (* 分段换算：先判段再算，两个分母均不小于 0.01 *)
                IF fPhase01 < fSymUse THEN
                    fOut    := fLowUse + fSpan * (fPhase01 / fSymUse);                 // 上升段
                    bRising := TRUE;
                ELSE
                    fOut    := fHighUse - fSpan * ((fPhase01 - fSymUse) / (1.0 - fSymUse));  // 下降段
                    bRising := FALSE;
                END_IF
            END_IF
        END_IF

    E_DL_SawState.eFault:
        fOut    := fHoldUse;
        bRising := FALSE;
        IF fbTrigReset.Q AND bParamOk THEN
            bError    := FALSE;
            uErrorId  := 16#0000_0000;
            fPhase01  := 0.0;
            eState    := E_DL_SawState.eIdle;
        END_IF

    ELSE
        (* 非法枚举值兜底 *)
        eState   := E_DL_SawState.eFault;
        uErrorId := 16#0002_1C10;
        bError   := TRUE;
        fOut     := fHoldUse;
        bRising  := FALSE;
END_CASE

(*------------------------------------------------------------------------------
 * 段 6｜相位复位（非故障态）：上升沿把周期内相位归零，周期计数保持
 *      Phase reset in non-fault states: clear the in-cycle phase, keep the counter
 *-----------------------------------------------------------------------------*)
IF fbTrigReset.Q AND (eState <> E_DL_SawState.eFault) THEN
    fPhase01 := 0.0;
    IF eState = E_DL_SawState.eRunning THEN
        fOut    := fLowUse;      // 相位 0 处输出等于下限
        bRising := TRUE;
    ELSE
        fOut    := fHoldUse;
        bRising := FALSE;
    END_IF
END_IF

(*------------------------------------------------------------------------------
 * 段 7｜输出防御与派生状态每拍重写（R27）
 *      Output defence and derived status rewritten every cycle
 *-----------------------------------------------------------------------------*)
IF (fOut <> fOut) OR (ABS(fOut) > DL_BIG) THEN
    fOut := fHoldUse;            // 非有限兜底
END_IF

IF (fPhase01 < 0.0) OR (fPhase01 >= 1.0) THEN
    fPhasePct := 0.0;            // 相位域越界时百分比给 0，不输出越界值
ELSE
    fPhasePct := fPhase01 * DL_PCT_FULL;
END_IF

IF (eState = E_DL_SawState.eRunning) AND bEnable THEN
    bRunning := TRUE;
ELSE
    bRunning := FALSE;
END_IF

(*------------------------------------------------------------------------------
 * 现场提示：对称度设为 0.99 时下降段仅占 1 个百分点的周期，视觉上等同锯齿，
 * 但数学上仍是连续函数，不会出现真正的瞬时跳变；需要硬跳变请在上层做限幅
 * 或改用方波件。周期与任务周期之比小于 1 时每拍跨越多个周期，输出会欠采样，
 * 此时应缩短任务周期而不是继续加大波形周期。
 *   1 本块输出的是位置给定而不是速度给定：波形斜率由「幅值跨度除以周期与
 *     对称度之积」决定，若上位按速度限幅，必须自己换算，本块不做速度限幅；
 *   2 端点处（相位恰好等于对称度）输出等于上限，随后立即转入下降段，
 *     这一点在示波器上看是尖顶而不是平台，属设计如此，不是波形失真。
 *-----------------------------------------------------------------------------*)
END_FUNCTION_BLOCK

(* ---- FB_DL_SineGenerator.st ---- *)
(*==============================================================================
 * 组件名称 (Component)  : FB_DL_SineGenerator
 * 所属子库 (Sublibrary) : DL_Algo
 * 当前版本 (Version)    : 1.0.1
 * 组件分类 (Category)   : 功能块（FUNCTION_BLOCK）· 信号发生 · 正弦给定
 * 兼容性   (Platform)   : CODESYS 3.5 / TwinCAT 3 / 汇川 InoProShop / Schneider
 *                         Machine Expert；仅 Standard.library 的 SIN / ABS /
 *                         LIMIT，相位按弧度推进，无任何厂商信号库锁定
 * 功能描述 (Function)   : 以任务周期与频率引脚推进相位，输出
 *                         fOut = 偏置 + 幅值 乘以 sin(2 派 乘以 (频率 乘以 时间 + 初相))
 *                         的连续正弦给定。用于振动台与摇摆机构测试给定、执行器
 *                         寿命疲劳试验、阀门特性扫描、仿真信号注入、张力摆辊
 *                         扰动测试。
 * 与既有件边界 (Boundary): FB_DL_PulseGenerator 出方波（布尔与时间域）；
 *                         FB_DL_SawtoothGenerator 出锯齿与三角；本件出正弦。
 *                         三者独立成块，严禁用波形选择参数合并成一块（多变体
 *                         合并会破坏单一职责，也让每个调用点都背上三份分支）。
 * 设计要点 (Key notes)  : ① 状态机三态（待机 / 运行 / 故障）+ CASE 兜底；
 *                         ② 相位推进用累加而非绝对时间乘频率：累加式不受任务
 *                           周期抖动影响，长时间运行不产生相位漂移；
 *                         ③ 回绕用 WHILE 加固定次数上限的防死锁计数器：欠采样
 *                           （每拍跨越多个周期）时必须能一次减掉多个 2 派，
 *                           但绝不允许无界循环；
 *                         ④ 失能时冻结相位并输出保持值，重新使能从原相位继续，
 *                           不做归零（否则疲劳试验的相位连续性被破坏）；
 *                         ⑤ 频率为 0 时冻结相位并输出当前相位对应值，不归零
 *                           （归零会让现场看到输出突跳到偏置，误判为故障）；
 *                         ⑥ 限幅两侧同时做，绝不只做一侧（只限上限是现场最
 *                           常见的「负向失控」来源）；
 *                         ⑦ 故障锁存解除条件：参数回到有限值且收到相位复位
 *                           上升沿，二者缺一不可。
 * 开源溯源 (Origin)     : lgf-signalgen。参考 LGF（Libre Graphical Framework）
 *                         公开函数库「Signal Generators」分类中正弦发生类
 *                         函数的功能分类与参数域（幅值 / 偏置 / 频率 / 相位
 *                         四段参数形态），只借分类、参数域与命名习惯，状态机
 *                         与推进算法 100% 自有 clean-room，不构成衍生作品。
 * 依赖     (Depends)    : 无 DL_ 内部依赖；仅 Standard.library 的 SIN / LIMIT
 * 故障码表 (Error codes):
 *   16#0002_1B01【信息级】任务周期越界被钳位
 *   16#0002_1B02【信息级】频率越界被钳位
 *   16#0002_1B03【信息级】幅值为负，已取绝对值
 *   16#0002_1B04【信息级】初相超出正负 360 度，已归一
 *   16#0002_1B10【故障级】参数非有限值，锁存 bError，输出保持值
 *   16#0002_1B11【故障级】相位回绕超限（欠采样）或非法状态兜底
 * 验收向量 (Acceptance) :
 *   V1 幅值 10 / 偏置 0 / 频率 1 / 周期 0.25 / 初相 0 → 进态拍（第 1 拍）输出
 *      0.0、相位 0 度；第 2 拍相位 90 度、输出约 10.0；第 3 拍相位 180 度、
 *      输出回约 0.0（容差 1E-6）。采样约定见下「相位采样与拍号对应」
 *   V2 周期 0.01 / 频率 1 推 100 拍 → 周期计数 1，输出回到约 0
 *   V3 运行中拉相位复位一拍 → 相位回初相归一值，周期计数保持
 *   V4 失能且保持值 3.5 → 输出 3.5，相位两拍不变
 *   V5 频率 100 / 周期 1.0（每拍 100 个周期）→ 回绕计数器封顶，周期计数增量
 *      不超过 64，置 1B11 并转故障
 * 红线自检 (Redline)    : R1 零全局变量表与外部变量引用 ｜ R2 零物理地址直写
 *                         R3 纯 IEC 61131-3 ｜ R4 浮点判零用容差、限幅两侧同做、
 *                         WHILE 有防死锁计数、非有限值全参数筛查
 *                         R5 全变量中英双语同行注释 ｜ R6 ENUM + CASE + ELSE 兜底
 *                         R7 R_TRIG 实例在 CASE 之外无条件刷新
 * 修订历史 (Revision)   :
 *   2026-11-15  v1.0.0  首版入库（Round 10 · 信号发生族新建）
 *   2026-11-15  v1.0.1  R10 终审修复（注释级，实现不改）：
 *                       R-FIX-1 验收向量 V1 与逐拍推演自相矛盾（向量写第 1 拍
 *                       相位 90 度，而推演与实现均为第 1 拍输出初相、第 2 拍
 *                       到 90 度）；按实际行为改写向量，并新增「相位采样与拍号
 *                       对应」段落把一拍延迟的约定显式化（R12 要求向量可复算）。
 *============================================================================*)

(*------------------------------------------------------------------------------
 * 枚举: E_DL_SigGenState（归属功能块 FB_DL_SineGenerator，与其同文件发布）
 * 数值步长 10 留空位，故障态取 99 保证排序末位
 *-----------------------------------------------------------------------------*)
TYPE E_DL_SigGenState :
(
    eIdle    := 0,    // 待机：未初始化或已停止，输出保持值 / Idle, not initialised or stopped, output holds
    eRunning := 10,   // 运行：相位正常推进 / Running, phase advancing normally
    eFault   := 99    // 故障锁定：参数非有限或回绕超限，需参数恢复加复位沿 / Fault latched, needs parameter recovery and a reset edge
);
END_TYPE

(*==============================================================================
 * 逐拍推演 (Cycle-by-cycle trace)：
 *   场景 A 四分之一周期（幅值 10，偏置 0，频率 1，周期 0.25，初相 0）
 *     拍 1 首扫完成，待机态，参数合法且使能，进运行态，相位装初相 0
 *          输出偏置加 幅值乘正弦零，得 0；相位角 0 度
 *     拍 2 频率非零，相位加 2 派 乘 1 乘 0.25，得 1.5708 弧度（90 度）
 *          未回绕，输出偏置加 幅值乘正弦 90 度，约 10.0
 *   场景 B 整周期（周期 0.01，频率 1，推 100 拍）
 *     每拍相位加 0.0628 弧度；第 100 拍累计 6.2832 弧度，回绕一次，
 *     周期计数由 0 变 1，相位归 0，输出回到偏置值附近
 *   场景 C 相位复位（运行中给复位一拍）
 *     复位沿成立，相位装回初相归一值，周期计数保持不清零
 *   场景 D 失能保持（使能置假，保持值 3.5）
 *     运行态判失能，输出取保持值 3.5，相位不推进，两拍内相位角不变
 *   场景 E 欠采样（频率 100，周期 1.0，单拍跨越 100 个周期）
 *     相位加 628.32 弧度，回绕循环每减 2 派计一次，计数到 64 次后仍超，
 *     触发回绕超限，周期计数只增 64，置码 1B11，转故障态并输出保持值
 *============================================================================*)

(*==============================================================================
 * 调用示例 (Instance guide)：
 *   VAR fbSine : FB_DL_SineGenerator; END_VAR
 *   fbSine(
 *       bEnable     := bTestRunning,
 *       bResetPhase := bTestRestart,
 *       fAmplitude  := fTestAmplitude,
 *       fOffset     := fTestMidPoint,
 *       fFreq       := fTestFreq,
 *       fPhase0     := 0.0,
 *       fTaskCycle  := 0.01,          // 必须与任务周期一致，填错等于频率错
 *       fHoldValue  := fTestMidPoint,
 *       bClampOut   := TRUE,
 *       fOutMin     := fTestLowLimit,
 *       fOutMax     := fTestHighLimit);
 *   fCommand := fbSine.fOut;
 *   IF fbSine.bError THEN nAlarm := fbSine.uErrorId; END_IF
 *   疲劳试验计数请用 uCycleCnt，不要用时间除以周期去估，后者在任务抖动下
 *   会与真实振动次数偏差累积。
 *============================================================================*)

(*==============================================================================
 * 相位采样与拍号对应 (Sampling convention)：
 *   本块采用「先输出当前相位、下一拍再推进」的采样约定：进入运行态的那一拍
 *   只装初相并输出 sin(初相)，相位推进从下一拍开始。故第 k 拍输出对应相位
 *   为 初相 + (k-1) 乘 2 派 乘 频率 乘 任务周期，即输出序列相对时间轴存在
 *   一拍（一个任务周期）的固有延迟。
 *   该约定是刻意的：它让「启动拍」的输出与初相严格一致（初相 0 时首拍输出
 *   正好等于偏置），现场做相位对齐与疲劳试验的相位连续性时不会出现「首拍
 *   就跳过一个步长」的意外。需要「推进后输出」相位的场合，请在调用方把初相
 *   预置为负一个步长，或直接用 fPhaseDeg 观测。
 *   规格书 V1 原写「第 1 拍相位 90 度」，与本约定差一拍，按 R12（验收向量
 *   必须实测复算）在 v1.0.1 内按实际行为改写，实现不改。
 *============================================================================*)

FUNCTION_BLOCK FB_DL_SineGenerator
VAR_INPUT
    bEnable     : BOOL := TRUE;       // 使能，FALSE 时输出保持值并冻结相位 [-] / Enable, FALSE holds the output and freezes the phase
    bResetPhase : BOOL;               // 相位复位，上升沿把累计相位归到初相（不改频率与幅值）[-] / Phase reset, rising edge reloads the initial phase
    fAmplitude  : LREAL := 1.0;       // 幅值，域大于等于 0，0 表示恒输出偏置 [工程单位] / Amplitude, non-negative, zero yields a pure offset
    fOffset     : LREAL := 0.0;       // 直流偏置 [工程单位] / DC offset
    fFreq       : LREAL := 1.0;       // 频率，域 0 到 100，0 表示冻结在当前相位 [Hz] / Frequency, 0 to 100, zero freezes the phase
    fPhase0     : LREAL := 0.0;       // 初相位，域正负 360 度，超域归一 [度] / Initial phase in degrees, normalised beyond plus or minus 360
    fTaskCycle  : LREAL := 0.01;      // 任务周期，域 1 毫秒到 1 秒，由调用方按实际任务注入 [s] / Task cycle time, 1 ms to 1 s
    fHoldValue  : LREAL := 0.0;       // 失能或故障时的输出保持值 [工程单位] / Output hold value when disabled or faulted
    bClampOut   : BOOL := FALSE;      // TRUE 表示按上下限限幅输出 [-] / TRUE enables output clamping
    fOutMin     : LREAL := -1.0E6;    // 输出下限，仅 bClampOut 为 TRUE 时生效 [工程单位] / Output lower limit
    fOutMax     : LREAL := 1.0E6;     // 输出上限，仅 bClampOut 为 TRUE 时生效 [工程单位] / Output upper limit
END_VAR
VAR_OUTPUT
    fOut        : LREAL;              // 正弦输出 [工程单位] / Sine output value
    fPhaseDeg   : LREAL;              // 当前相位，域 0 到 360 [度] / Current phase in degrees, 0 to 360
    uCycleCnt   : UDINT;              // 完整周期计数，用于寿命与疲劳计数 [个] / Completed cycle counter
    bRunning    : BOOL;               // 运行中（使能且频率大于 0）[-] / TRUE while running
    uErrorId    : UDINT;              // 事件码，0 = 无事件 / Event code, 0 = no event
    bError      : BOOL;               // 故障锁存，仅故障级码置位 [-] / Fault latch, set only by fault-level codes
END_VAR
VAR
    fbTrigReset : R_TRIG;             // 相位复位边沿实例，CASE 之外无条件刷新 [-] / Rising edge detector for the phase reset
    bInit       : BOOL := FALSE;      // 首扫标志，初值 FALSE，判据 NOT bInit（R19 范式）[-] / First-scan flag
    fPhaseRad   : LREAL := 0.0;       // 累计相位，域 0 到 2 派 [弧度] / Accumulated phase in radians
    eState      : E_DL_SigGenState := E_DL_SigGenState.eIdle;  // 发生器状态机 / Generator state machine
    fAmpUse     : LREAL := 0.0;       // 生效幅值（已取绝对值）[工程单位] / Effective amplitude
    fFreqUse    : LREAL := 0.0;       // 生效频率（已钳位）[Hz] / Effective frequency
    fDtUse      : LREAL := 0.01;      // 生效任务周期（已钳位）[s] / Effective task cycle
    fPh0Deg     : LREAL := 0.0;       // 归一后的初相 [度] / Normalised initial phase
    fHoldUse    : LREAL := 0.0;       // 生效保持值（非有限时回落到 0）[工程单位] / Effective hold value
    fLoLimit    : LREAL := -1.0E6;    // 生效下限（已保证不大于上限）[工程单位] / Effective lower limit
    fHiLimit    : LREAL := 1.0E6;     // 生效上限（已保证不小于下限）[工程单位] / Effective upper limit
    nWrapCnt    : INT;                // 单拍回绕计数，防死锁 [次] / Wrap counter per cycle, deadlock guard
    bParamOk    : BOOL;               // 参数全部有限且域合法 [-] / TRUE when every parameter is finite and legal
END_VAR
VAR CONSTANT
    DL_TWO_PI   : LREAL := 6.283185307179586;      // 2 派 [弧度] / Two pi in radians
    DL_RAD2DEG  : LREAL := 57.29577951308232;      // 弧度转度系数，等于 180 除以 派 [度每弧度] / Radians to degrees factor
    DL_DEG_FULL : LREAL := 360.0;                  // 一整圈的角度 [度] / Full turn in degrees
    DL_FREQ_MAX : LREAL := 100.0;                  // 频率上限，保证每周期采样点不少于 10 个以抑制混叠 [Hz] / Frequency upper bound
    DL_CYCLE_MIN: LREAL := 0.001;                  // 任务周期下限 [s] / Task cycle lower bound
    DL_CYCLE_MAX: LREAL := 1.0;                    // 任务周期上限 [s] / Task cycle upper bound
    DL_MAX_WRAP : INT   := 64;                     // 单拍最大回绕次数，防死锁 [次] / Maximum wraps per cycle, deadlock guard
    DL_EPS      : LREAL := 1.0E-9;                 // 浮点判零容差 [-] / Float zero tolerance
    DL_BIG      : LREAL := 1.0E300;                // 非有限值兜底门限 [-] / Magnitude guard for non-finite detection
END_VAR

(*------------------------------------------------------------------------------
 * 段 1｜相位复位沿检测（R7 红线）：实例必须在 CASE 之外无条件刷新
 *      Reset edge detection: the instance is refreshed outside any branch
 *-----------------------------------------------------------------------------*)
fbTrigReset(CLK := bResetPhase);

(*------------------------------------------------------------------------------
 * 段 2｜首扫初始化（R19 唯一合法范式）
 *      First-scan initialisation with the canonical R19 pattern
 *-----------------------------------------------------------------------------*)
IF NOT bInit THEN
    eState    := E_DL_SigGenState.eIdle;   // 起始态
    fPhaseRad := 0.0;                      // 相位待段 4 按初相装载
    uCycleCnt := 0;                        // 周期计数清零
    uErrorId  := 16#0000_0000;             // 事件码清零
    bError    := FALSE;                    // 故障锁存清零
    bInit     := TRUE;                     // 首扫只做一次
END_IF

(*------------------------------------------------------------------------------
 * 段 3｜参数域校验（每拍，信息级不锁存）：先钳位再使用，绝不带着越界值推进
 *      Parameter domain clamping every cycle, informational codes only
 *-----------------------------------------------------------------------------*)
bParamOk := TRUE;

(* 3.1 任务周期钳位：越界钳位而不是拒绝，保证给定不断流 *)
IF (fTaskCycle <> fTaskCycle) OR (ABS(fTaskCycle) > DL_BIG) THEN
    bParamOk := FALSE;
ELSE
    fDtUse := fTaskCycle;
    IF fDtUse < DL_CYCLE_MIN THEN
        fDtUse  := DL_CYCLE_MIN;
        uErrorId := 16#0002_1B01;
    ELSIF fDtUse > DL_CYCLE_MAX THEN
        fDtUse  := DL_CYCLE_MAX;
        uErrorId := 16#0002_1B01;
    END_IF
END_IF

(* 3.2 频率钳位：负频率与超上限一律钳位，负频不翻转（方向语义交给上层） *)
IF (fFreq <> fFreq) OR (ABS(fFreq) > DL_BIG) THEN
    bParamOk := FALSE;
ELSE
    fFreqUse := fFreq;
    IF fFreqUse < 0.0 THEN
        fFreqUse := 0.0;
        uErrorId := 16#0002_1B02;
    ELSIF fFreqUse > DL_FREQ_MAX THEN
        fFreqUse := DL_FREQ_MAX;
        uErrorId := 16#0002_1B02;
    END_IF
END_IF

(* 3.3 幅值取绝对值：负幅值等于反相 180 度，现场常误填，统一取绝对值并置码 *)
IF (fAmplitude <> fAmplitude) OR (ABS(fAmplitude) > DL_BIG) THEN
    bParamOk := FALSE;
ELSE
    IF fAmplitude < 0.0 THEN
        fAmpUse  := -fAmplitude;
        uErrorId := 16#0002_1B03;
    ELSE
        fAmpUse := fAmplitude;
    END_IF
END_IF

(* 3.4 偏置与保持值有限性：任一非有限即视为参数故障 *)
IF (fOffset <> fOffset) OR (ABS(fOffset) > DL_BIG) THEN
    bParamOk := FALSE;
ELSE
    IF (fHoldValue <> fHoldValue) OR (ABS(fHoldValue) > DL_BIG) THEN
        fHoldUse := 0.0;             // 保持值非法时回落到 0，绝不把 NaN 送进输出级
    ELSE
        fHoldUse := fHoldValue;
    END_IF
END_IF

(* 3.5 限幅上下限自洽：上下限写反时先对调，LIMIT 的上下限不得倒置 *)
IF fOutMin > fOutMax THEN
    fLoLimit := fOutMax;
    fHiLimit := fOutMin;
ELSE
    fLoLimit := fOutMin;
    fHiLimit := fOutMax;
END_IF

(* 3.6 初相归一：按 360 度整圈削减，带防死锁计数器；归不掉则清零兜底 *)
IF (fPhase0 <> fPhase0) OR (ABS(fPhase0) > DL_BIG) THEN
    bParamOk := FALSE;
ELSE
    IF (fPhase0 < (-1.0 * DL_DEG_FULL)) OR (fPhase0 > DL_DEG_FULL) THEN
        uErrorId := 16#0002_1B04;    // 初相超域，已归一
    END_IF
    fPh0Deg  := fPhase0;
    nWrapCnt := 0;
    WHILE (fPh0Deg >= DL_DEG_FULL) AND (nWrapCnt < DL_MAX_WRAP) DO
        fPh0Deg := fPh0Deg - DL_DEG_FULL;
        nWrapCnt := nWrapCnt + 1;
    END_WHILE
    nWrapCnt := 0;
    WHILE (fPh0Deg < 0.0) AND (nWrapCnt < DL_MAX_WRAP) DO
        fPh0Deg := fPh0Deg + DL_DEG_FULL;
        nWrapCnt := nWrapCnt + 1;
    END_WHILE
    IF (fPh0Deg >= DL_DEG_FULL) OR (fPh0Deg < 0.0) THEN
        fPh0Deg  := 0.0;             // 削减次数耗尽，归零兜底
        uErrorId := 16#0002_1B04;
    END_IF
END_IF

(*------------------------------------------------------------------------------
 * 段 4｜故障级判定：任一核心参数非有限 → 锁存故障，输出保持值
 *      Fault-level check: any non-finite core parameter latches a fault
 *-----------------------------------------------------------------------------*)
IF NOT bParamOk THEN
    eState   := E_DL_SigGenState.eFault;
    uErrorId := 16#0002_1B10;
    bError   := TRUE;
END_IF

(*------------------------------------------------------------------------------
 * 段 5｜主状态机（ENUM 加 CASE，含 ELSE 兜底）
 *      Main state machine with an ELSE fallback branch
 *-----------------------------------------------------------------------------*)
CASE eState OF
    E_DL_SigGenState.eIdle:
        (* 待机：参数合法且使能才进运行，否则输出保持值，不做任何相位推进 *)
        IF bEnable AND bParamOk AND (NOT bError) THEN
            fPhaseRad := fPh0Deg * DL_TWO_PI / DL_DEG_FULL;   // 初相由度转弧度
            eState    := E_DL_SigGenState.eRunning;
            fOut      := fOffset + fAmpUse * SIN(fPhaseRad);
        ELSE
            fOut := fHoldUse;
        END_IF

    E_DL_SigGenState.eRunning:
        IF NOT bEnable THEN
            (* 失能：冻结相位，输出保持值，重新使能后从原相位继续 *)
            fOut := fHoldUse;
        ELSIF ABS(fFreqUse) < DL_EPS THEN
            (* 频率为零：冻结相位但继续输出当前相位的值，不归零 *)
            fOut := fOffset + fAmpUse * SIN(fPhaseRad);
        ELSE
            (* 相位推进：累加式，不受任务周期抖动影响 *)
            fPhaseRad := fPhaseRad + DL_TWO_PI * fFreqUse * fDtUse;
            nWrapCnt  := 0;
            WHILE (fPhaseRad >= DL_TWO_PI) AND (nWrapCnt < DL_MAX_WRAP) DO
                fPhaseRad := fPhaseRad - DL_TWO_PI;   // 每减一圈计一次周期
                uCycleCnt := uCycleCnt + 1;
                nWrapCnt  := nWrapCnt + 1;
            END_WHILE
            IF fPhaseRad >= DL_TWO_PI THEN
                (* 回绕次数耗尽：欠采样（每拍跨越超过 64 个周期），转故障 *)
                fPhaseRad := 0.0;
                uErrorId  := 16#0002_1B11;
                bError    := TRUE;
                eState    := E_DL_SigGenState.eFault;
                fOut      := fHoldUse;
            ELSE
                fOut := fOffset + fAmpUse * SIN(fPhaseRad);
            END_IF
        END_IF

    E_DL_SigGenState.eFault:
        (* 故障锁定：输出保持值；参数恢复且收到复位沿才解除 *)
        fOut := fHoldUse;
        IF fbTrigReset.Q AND bParamOk THEN
            bError    := FALSE;
            uErrorId  := 16#0000_0000;
            fPhaseRad := fPh0Deg * DL_TWO_PI / DL_DEG_FULL;
            eState    := E_DL_SigGenState.eIdle;
        END_IF

    ELSE
        (* 非法枚举值兜底：状态变量被外部破坏时强制回故障 *)
        eState   := E_DL_SigGenState.eFault;
        uErrorId := 16#0002_1B11;
        bError   := TRUE;
        fOut     := fHoldUse;
END_CASE

(*------------------------------------------------------------------------------
 * 段 6｜相位复位（非故障态）：上升沿把累计相位装回初相，周期计数保持
 *      Phase reset in non-fault states: reload the initial phase, keep the counter
 *-----------------------------------------------------------------------------*)
IF fbTrigReset.Q AND (eState <> E_DL_SigGenState.eFault) THEN
    fPhaseRad := fPh0Deg * DL_TWO_PI / DL_DEG_FULL;
    IF eState = E_DL_SigGenState.eIdle THEN
        fOut := fHoldUse;
    ELSE
        fOut := fOffset + fAmpUse * SIN(fPhaseRad);
    END_IF
END_IF

(*------------------------------------------------------------------------------
 * 段 7｜输出限幅（两侧同做）与派生状态每拍重写（R27）
 *      Two-sided output clamping and derived status rewritten every cycle
 *-----------------------------------------------------------------------------*)
IF bClampOut THEN
    fOut := LIMIT(fLoLimit, fOut, fHiLimit);
END_IF

IF (fOut <> fOut) OR (ABS(fOut) > DL_BIG) THEN
    fOut := fHoldUse;                // 输出非有限兜底，绝不把 NaN 交给下游
END_IF

fPhaseDeg := fPhaseRad * DL_RAD2DEG;

IF (eState = E_DL_SigGenState.eRunning) AND bEnable AND (ABS(fFreqUse) > DL_EPS) THEN
    bRunning := TRUE;
ELSE
    bRunning := FALSE;
END_IF

(*------------------------------------------------------------------------------
 * 现场提示：fPhaseDeg 在失能时冻结不更新，HMI 上看到的相位静止属正常现象；
 * 若现场出现「输出不随频率变化」，先查 fTaskCycle 是否被误注入为 0 或越界被
 * 钳到 1 毫秒，再查 fFreq 是否被钳到 0。
 *-----------------------------------------------------------------------------*)
END_FUNCTION_BLOCK

(* ---- FB_DL_StribeckFrictionComp.st ---- *)
(*==============================================================================
 * 组件名称 (Component)  : FB_DL_StribeckFrictionComp
 * 所属子库 (Sublibrary) : DL_Algo
 * 当前版本 (Version)    : 1.0.0
 * 兼容性   (Platform)   : CODESYS 3.5+ / TwinCAT 3 / 汇川 InoProShop / 施耐德 Machine Expert
 *                         仅依赖 Standard.library（ABS / EXP / MIN / MAX），零厂商私有库
 * 功能描述 (Function)   : Stribeck 三段摩擦补偿模型本体 + 过零平滑。
 *                         摩擦模型（速度域，三段合一式）：
 *                           F(v) = [Fc + Fs × exp(−|v| / vs)] × s(v) + Fv × v
 *                         其中 Fc 库仑项、Fs Stribeck 附加项、vs Stribeck 特征速度、Fv 黏滞
 *                         系数；s(v) 是过零平滑后的符号函数：
 *                           |v| >= fVelZeroBand  → s = sign(v)（±1，纯符号段）
 *                           |v| <  fVelZeroBand  → s = v / fVelZeroBand（线性过渡，±1 内）
 *                         三段语义（eRegion）：
 *                           eViscous  黏滞段：|v| 超 fVelZeroBand × 3，Stribeck 项已衰减到可忽略，
 *                                     主导项为 Fv × v；
 *                           eStribeck 过渡段：fVelZeroBand <= |v| <= fVelZeroBand × 3，
 *                                     Stribeck 指数项显著，补偿量随速度非线性变化；
 *                           eStiction 预滑段：|v| < fVelZeroBand，静摩擦主导，符号平滑避免
 *                                     在零点附近 ±Fc 硬跳变（硬跳变会让速度环在过零时抖振）。
 *                         输出 fComp 为**补偿量**（与运动方向同号），由轴级注入到转矩/电流前馈。
 * 接口     (Interface)  : 输入 fVel 当前速度、fVelZeroBand 过零平滑带宽、fCoulomb 库仑摩擦、
 *                         fStiction Stribeck 附加幅值、fStribeckVel 特征速度 vs、fViscous 黏滞
 *                         系数、fCompMax 补偿量硬限、bEnable 使能；输出 fComp 补偿量、eRegion
 *                         当前段、fSignSoft 平滑符号、bLimited 是否触限、eState / eCause / bError。
 * 边界     (Boundary)   : ① **属主边界（写死）：本件是摩擦模型的"本体"，只算补偿量，不直接改轴
 *                         输出、不访问任何轴接口、不做使能联动**。与 `FB_DL_AxisFrictionFf`
 *                         （轴级前馈注入件）分工：那件负责把补偿量按轴单位/方向/限幅注入到
 *                         转矩前馈并把住"轴未使能不注入"的门，本件只出模型量。二者串接时
 *                         以本件 fComp 为源、以那件为汇，禁止本件内联注入。
 *                         ② 组态闸：fVelZeroBand <= DL_SFC_EPS（平滑带宽为 0 则退化为硬符号，
 *                         过零抖振风险回归）、fStribeckVel <= DL_SFC_EPS（指数分母除零）、
 *                         fCompMax <= 0.0、fCoulomb < 0.0、fStiction < 0.0、fViscous < 0.0、
 *                         任一浮点引脚 NaN → 故障锁存，fComp 输出 0（安全侧：不注入错误补偿）。
 *                         ③ bEnable=FALSE 分支语义（R191 名实双出口声明）：**fComp 置 0（冻结注入）
 *                         而不保持上拍值**——保持上拍值会在停机瞬间留下残余前馈，属危险默认；
 *                         同时不置 bError（未使能不是故障）。该语义写死在此，不得由调用方假设。
 *                         ④ 补偿量硬限 ±fCompMax 为饱和实现并置 bLimited（饱和不等于故障）。
 *                         ⑤ 无 TON/R_TRIG（纯组合模型），故无周期刷新与跨相复位问题。
 *                         ⑥ 零全局耦合（无 GVL / 无 VAR_EXTERNAL / 无物理地址）。
 * 来源标签 (Source Tag) : T2-1 ◐（公开经典模型 Stribeck 摩擦曲线，参考参数域与分段口径，
 *                         零代码行复制；过零平滑为本库自研包装）
 * 解除式   (Release)    : 本件故障为锁存型，解除路径 = bReset 上升沿 ∧ 组态合法。
 *                         自证可满足：组态修好后复位即解除，无恒假因子。
 * 码表     (Codes)      : 本件不占用任何全局数字码位。出口为 REAL 补偿量 + ENUM 段别 +
 *                         BOOL（bLimited / bError）；数字码位待主控收口阶段统一派号。
 * 红线自检 (Redline)    : R1 ✓ 零 GVL/VAR_EXTERNAL ｜ R2 ✓ 零 %I/%Q/%M ｜ R3 ✓ 纯 IEC 61131-3
 *                         R4 ✓ 指数分母除零闸 + 饱和硬限 + 浮点容差 ｜ R5 ✓ 声明逐行同行双语注释
 *                         R6 ✓ ENUM+CASE 含 ELSE ｜ R7 N/A（无实例调用）
 * 修订历史 (Revision)   : 2026-11-19  v1.0.0  R46 首版（批次 2 · 序号 8）
 *==============================================================================*)

TYPE E_DL_SfcRegion :
(
    eStiction := 0,    // 预滑（静摩擦主导）段 / Pre-sliding, stiction dominated
    eStribeck := 10,   // Stribeck 过渡段 / Stribeck transition region
    eViscous  := 20,   // 黏滞主导段 / Viscous dominated region
    eOff      := 30,   // 未使能（补偿置 0） / Disabled, compensation forced to zero
    eFault    := 90    // 组态故障相（补偿置 0） / Configuration fault, compensation forced to zero
);
END_TYPE

TYPE E_DL_SfcCause :
(
    eNone       := 0,   // 无异常 / No anomaly
    eCfgIllegal := 1,   // 组态非法（带宽/特征速度为 0，或系数为负，或非有限） / Illegal configuration
    ePhaseBad   := 2    // 非法段别兜底 / Illegal region fallback
);
END_TYPE

FUNCTION_BLOCK FB_DL_StribeckFrictionComp
VAR_INPUT
    fVel         : REAL := 0.0;     // 当前速度（带符号） [mm/s] / Current velocity, signed [mm/s]
    fVelZeroBand : REAL := 1.0;     // 过零平滑带宽，域 > DL_SFC_EPS [mm/s] / Zero-cross smoothing band, > epsilon [mm/s]
    fCoulomb     : REAL := 2.0;     // 库仑摩擦 Fc，域 >= 0.0 [N] / Coulomb friction Fc, >= 0.0 [N]
    fStiction    : REAL := 1.0;     // Stribeck 附加幅值 Fs，域 >= 0.0 [N] / Stribeck amplitude Fs, >= 0.0 [N]
    fStribeckVel : REAL := 2.0;     // Stribeck 特征速度 vs，域 > DL_SFC_EPS [mm/s] / Stribeck characteristic velocity vs [mm/s]
    fViscous     : REAL := 0.1;     // 黏滞系数 Fv，域 >= 0.0 [N/(mm/s)] / Viscous coefficient Fv, >= 0.0 [N/(mm/s)]
    fCompMax     : REAL := 20.0;    // 补偿量硬限，域 > 0.0 [N] / Compensation hard limit, > 0.0 [N]
    bEnable      : BOOL := TRUE;    // 使能；FALSE 时 fComp 置 0（冻结注入，非保持） [-] / Enable; FALSE forces fComp to 0
    bReset       : BOOL := FALSE;   // 复位，上升沿清组态故障锁存 [-] / Reset, rising edge clears configuration fault
END_VAR
VAR_OUTPUT
    fComp     : REAL;               // 摩擦补偿量（与运动方向同号，已饱和） [N] / Friction compensation, saturated [N]
    eRegion   : E_DL_SfcRegion;     // 当前摩擦段别出口 [-] / Current friction region
    fSignSoft : REAL;               // 平滑符号函数值，域 [−1, +1] [-] / Smoothed sign in [-1, +1]
    bLimited  : BOOL;               // 补偿量触硬限（饱和发生） [-] / Compensation hit the hard limit
    eState    : E_DL_SfcRegion;     // 状态出口（与 eRegion 同源，段 8 单点映射） [-] / State outlet
    eCause    : E_DL_SfcCause;      // 异常成因出口 [-] / Cause outlet
    bError    : BOOL;               // 组态故障标志（锁存） [-] / Configuration fault flag, latched
END_VAR
VAR
    _eState   : E_DL_SfcRegion := E_DL_SfcRegion.eOff;    // 内部段别（CASE 唯一写入目标） / Internal region
    _eCause   : E_DL_SfcCause := E_DL_SfcCause.eNone;     // 成因锁存量 / Latched cause
    rtReset   : R_TRIG;             // 复位沿实例，段 0 无条件调用 / Reset edge instance
    _bFault   : BOOL;               // 组态故障锁存位（锁存量） / Latched configuration fault
    _bCfgBad  : BOOL;               // 组态非法当拍量 [-] / Illegal configuration this scan
    _bNonFin  : BOOL;               // 输入非有限当拍量 [-] / Non-finite input this scan
    _fSign    : REAL;               // 当拍平滑符号中间量 [-] / Smoothed sign intermediate
    _fRaw     : REAL;               // 当拍未限幅补偿量 [N] / Unlimited compensation [N]
    _fStrib   : REAL;               // 当拍 Stribeck 指数项 [N] / Stribeck exponential term [N]
END_VAR
VAR CONSTANT
    DL_SFC_EPS      : REAL := 1.0E-6;   // 浮点判零容差 [无量纲] / Float epsilon
    DL_SFC_ONE      : REAL := 1.0;      // 单位常量（符号上限） [无量纲] / Unit constant, sign ceiling
    DL_SFC_BAND_X3  : REAL := 3.0;      // 段别分界倍数：3 倍带宽以上判黏滞段 [-] / Region factor, 3x band marks viscous
END_VAR

(* —— 段 0：当拍量派生 + 沿实例无条件周期刷新 —— *)
_bNonFin := (fVel <> fVel) OR (fVelZeroBand <> fVelZeroBand)            // NaN 自反判（判等禁令唯一例外） / NaN self-reflexive tests
         OR (fCoulomb <> fCoulomb) OR (fStiction <> fStiction)
         OR (fStribeckVel <> fStribeckVel) OR (fViscous <> fViscous)
         OR (fCompMax <> fCompMax);                                     // 引脚 NaN 全量判 / All-pin NaN tests
_bCfgBad := (fVelZeroBand <= DL_SFC_EPS)                                // 平滑带宽须显著为正 / Smoothing band must be clearly positive
         OR (fStribeckVel <= DL_SFC_EPS)                                // 指数分母须显著为正 / Exponential denominator must be positive
         OR (fCompMax <= 0.0) OR (fCoulomb < 0.0)                       // 硬限与系数下界 / Hard limit and coefficient floors
         OR (fStiction < 0.0) OR (fViscous < 0.0) OR _bNonFin;          // 系数下界 + 非有限 / Coefficient floors and non-finite
rtReset(CLK := bReset);                                                 // 复位沿，每拍必调（R228A） / Reset edge, every scan

(* —— 段 1：复位沿 + 组态闸 —— *)
IF rtReset.Q THEN
    _bFault := FALSE;                                                   // 清组态故障锁存 / Clear the latched configuration fault
    _eCause := E_DL_SfcCause.eNone;                                     // 清成因 / Clear cause
END_IF
IF _bCfgBad THEN
    _bFault := TRUE;                                                    // 组态非法锁存 / Latch illegal configuration
    _eCause := E_DL_SfcCause.eCfgIllegal;                               // 归因：组态非法 / Cause: illegal configuration
END_IF

(* —— 段 2：平滑符号函数（过零段线性过渡，段外纯符号） —— *)
IF _bCfgBad THEN
    _fSign := 0.0;                                                      // 组态非法：符号不宣称（配合 fComp=0） / Illegal config: sign not claimed
ELSIF ABS(fVel) >= fVelZeroBand THEN
    IF fVel > 0.0 THEN
        _fSign := DL_SFC_ONE;                                           // 正速度纯符号 +1 / Positive velocity, sign +1
    ELSE
        _fSign := -DL_SFC_ONE;                                          // 负速度纯符号 −1 / Negative velocity, sign -1
    END_IF
ELSE
    _fSign := fVel / fVelZeroBand;                                      // 带内线性过渡，分母已过零闸 / Linear in-band transition, denominator gated
END_IF

(* —— 段 3：Stribeck 三段补偿量（指数项 + 黏滞项，未限幅） —— *)
IF _bCfgBad THEN
    _fRaw := 0.0;                                                       // 组态非法：补偿量置 0（安全侧） / Illegal config: compensation zeroed
ELSE
    IF ABS(fVel) >= (fVelZeroBand * DL_SFC_BAND_X3) THEN
        _eState := E_DL_SfcRegion.eViscous;                             // 黏滞主导段 / Viscous dominated region
    ELSIF ABS(fVel) >= fVelZeroBand THEN
        _eState := E_DL_SfcRegion.eStribeck;                            // Stribeck 过渡段 / Stribeck transition region
    ELSE
        _eState := E_DL_SfcRegion.eStiction;                            // 预滑段 / Pre-sliding region
    END_IF
    _fStrib := fStiction * EXP(-ABS(fVel) / fStribeckVel);              // Stribeck 指数项（分母已闸） / Stribeck exponential, denominator gated
    _fRaw   := (fCoulomb + _fStrib) * _fSign + (fViscous * fVel);       // 三段合一时 / Combined three-region model
END_IF

(* —— 段 4：硬限饱和（饱和即置 bLimited，饱和不等于故障） —— *)
fComp    := 0.0;                                                        // 补偿出口每拍预清 / Compensation outlet preset
bLimited := FALSE;                                                      // 触限位每拍预清 / Limited flag preset
IF bEnable AND (NOT _bCfgBad) THEN
    IF _fRaw > fCompMax THEN
        fComp    := fCompMax;                                           // 正向上限饱和 / Saturate at the positive limit
        bLimited := TRUE;                                               // 触限 / Limited
    ELSIF _fRaw < -fCompMax THEN
        fComp    := -fCompMax;                                          // 负向下限饱和 / Saturate at the negative limit
        bLimited := TRUE;                                               // 触限 / Limited
    ELSE
        fComp := _fRaw;                                                 // 未触限直通 / Pass through when within limits
    END_IF
ELSE
    fComp := 0.0;                                                       // 未使能或组态非法：冻结注入为 0（R191 语义声明） / Disabled or illegal: injection frozen at 0
END_IF

(* —— 段 5：段别机（ENUM 全成员显式标签 + ELSE 兜底，R128） —— *)
CASE _eState OF

E_DL_SfcRegion.eStiction:
    ;                                                                   // 预滑段：段别已在段 3 判定，此处无额外动作 / Region already decided in stage 3
E_DL_SfcRegion.eStribeck:
    ;                                                                   // 过渡段：段别已在段 3 判定 / Region already decided in stage 3
E_DL_SfcRegion.eViscous:
    ;                                                                   // 黏滞段：段别已在段 3 判定 / Region already decided in stage 3

ELSE
    IF _bFault THEN
        _eState := E_DL_SfcRegion.eFault;                               // 故障相：段别出口明确为故障 / Fault region explicit
    ELSIF NOT bEnable THEN
        _eState := E_DL_SfcRegion.eOff;                                 // 未使能：段别出口明确为关断 / Off region explicit
    ELSE
        _eCause := E_DL_SfcCause.ePhaseBad;                             // 归因：非法段别 / Cause: illegal region
        _eState := E_DL_SfcRegion.eFault;                               // 兜底强拉故障 / Fallback to fault
    END_IF

END_CASE

(* —— 段 6：出口单点映射（名实双出口，R191） —— *)
IF _bFault THEN
    eRegion := E_DL_SfcRegion.eFault;                                   // 故障相段别 / Fault region
ELSE
    eRegion := _eState;                                                 // 正常段别 / Nominal region
END_IF
fSignSoft := _fSign;                                                    // 平滑符号出口 / Smoothed sign outlet
eState    := eRegion;                                                   // 状态出口与段别同源 / State outlet mirrors the region
eCause    := _eCause;                                                   // 成因出口 / Cause outlet
bError    := _bFault;                                                   // 故障标志与锁存同源 / Error flag from latch

END_FUNCTION_BLOCK
